{region 'Documentation'}
(*!
<summary>Checks results and isolated findings before allowing the script to advance.</summary>
*)
{endregion}
METHOD PROTECTED ProcessAssertions
VAR_INPUT
    Enable : BOOL; //! Phase permission supplied by the owning Test Case; FALSE does not authorize progression, while observation may continue.
END_VAR
VAR
    Evaluate : BOOL;
    FindingIndex : UINT;
    DetailsMatch : BOOL;
    FindingMatches : BOOL;
    ExpectedMessage : STRING(GVL_Constants.MessageLength);
END_VAR
FFirstCycleGate(Enable := Enable AND FGateObservationReady,
    State := State,
    IN := FGateMatches);
Evaluate := Enable AND FObservationReady;
FIsNaNResult(Enable := Evaluate,
    State := State,
    IN := FIsNaNSubject.Result = FExpectedIsNaN);
FIsFiniteResult(Enable := Evaluate,
    State := State,
    IN := FIsFiniteSubject.Result = FExpectedIsFinite);
FIsInfiniteResult(Enable := Evaluate,
    State := State,
    IN := FIsInfiniteSubject.Result = FExpectedIsInfinite);
DetailsMatch := TRUE;
FindingIndex := 1;
IF Evaluate THEN
    IF FFindingIsNaN <> E_Result.NotEvaluated THEN
        ExpectedMessage := CONCAT('Assertion failed: expected NaN. Actual = ',
            CreateAssertionTextValue_LReal(Value := FValue.Value));
        ExpectedMessage := CONCAT(ExpectedMessage, '.');
        FindingMatches := IsFindingValid(Index := FindingIndex,
            ExpectedName := FIsNaNSubject.Name,
            ExpectedResult := FFindingIsNaN,
            ExpectedMessage := ExpectedMessage);
        DetailsMatch := DetailsMatch AND FindingMatches;
        FindingIndex := FindingIndex + 1;
    END_IF;
    IF FFindingIsFinite <> E_Result.NotEvaluated THEN
        ExpectedMessage := CONCAT('Assertion failed: expected a finite value. Actual = ',
            CreateAssertionTextValue_LReal(Value := FValue.Value));
        ExpectedMessage := CONCAT(ExpectedMessage, '.');
        FindingMatches := IsFindingValid(Index := FindingIndex,
            ExpectedName := FIsFiniteSubject.Name,
            ExpectedResult := FFindingIsFinite,
            ExpectedMessage := ExpectedMessage);
        DetailsMatch := DetailsMatch AND FindingMatches;
        FindingIndex := FindingIndex + 1;
    END_IF;
    IF FFindingIsInfinite <> E_Result.NotEvaluated THEN
        ExpectedMessage := CONCAT('Assertion failed: expected positive or negative infinity. Actual = ',
            CreateAssertionTextValue_LReal(Value := FValue.Value));
        ExpectedMessage := CONCAT(ExpectedMessage, '.');
        FindingMatches := IsFindingValid(Index := FindingIndex,
            ExpectedName := FIsInfiniteSubject.Name,
            ExpectedResult := FFindingIsInfinite,
            ExpectedMessage := ExpectedMessage);
        DetailsMatch := DetailsMatch AND FindingMatches;
        FindingIndex := FindingIndex + 1;
    END_IF;
END_IF;
FCaptureIntegrity(Enable := Evaluate,
    State := State,
    IN := (FCaptureStatus.SequenceId = UINT_TO_UDINT(FindingIndex - 1))
        AND (FCaptureStatus.LostEventCount = 0)
        AND (FCaptureFifo.ElementCount = FindingIndex - 1));
FFindingDetails(Enable := Evaluate,
    State := State,
    IN := DetailsMatch);
IF Evaluate THEN
    FChecked := TRUE;
END_IF;
END_METHOD

{region 'Documentation'}
(*!
<summary>No Preparation phase is required.</summary>
*)
{endregion}
METHOD PROTECTED ProcessPreparations
VAR_INPUT
    // SA0033: Required hook; no Preparation phase.
    {attribute 'analysis' := '-33'}
    Enable : BOOL; //! Phase permission supplied by the owning Test Case; FALSE does not authorize progression, while observation may continue.
END_VAR
END_METHOD

{region 'Documentation'}
(*!
<summary>Restarts the row script and resets outer verdicts.</summary>
*)
{endregion}
METHOD PROTECTED ProcessReset
FFirstCycleGate.Reset();
FFirstCyclePending := FALSE;
FGateObservationReady := FALSE;
FGateMatches := FALSE;
FRow := RowQuietNaN;
FRowPrepared := FALSE;
FRepeatChecked := FALSE;
FChecked := FALSE;
FObservationReady := FALSE;
FIsNaNResult.Reset();
FIsFiniteResult.Reset();
FIsInfiniteResult.Reset();
FCaptureIntegrity.Reset();
FFindingDetails.Reset();
CompleteReset();
END_METHOD

{region 'Documentation'}
(*!
<summary>Prepares, checks and repeats each row over separate PLC cycles.</summary>
*)
{endregion}
METHOD PROTECTED ProcessTests
VAR_INPUT
    Enable : BOOL; //! Phase permission supplied by the owning Test Case; FALSE does not authorize progression, while observation may continue.
END_VAR
IF NOT Enable THEN
    RETURN;
END_IF;

FGateObservationReady := FALSE;
IF FChecked THEN
    FChecked := FALSE;
    FObservationReady := FALSE;
    IF FRepeatChecked THEN
        IF FRow = LastRow THEN
            CompleteTests();
            RETURN;
        END_IF;
        FRow := FRow + 1;
        FRowPrepared := FALSE;
        FRepeatChecked := FALSE;
    ELSE
        FRepeatChecked := TRUE;
    END_IF;
END_IF;

IF NOT FRowPrepared THEN
    SelectRow();
    FCapture.Reset();
    IF NOT FPreserveResults THEN
        ResetSubjects();
    END_IF;
    CallSubjects(Enable := FALSE);
    FRowPrepared := TRUE;
    FFirstCyclePending := TRUE;
ELSIF FFirstCyclePending THEN
    CallSubjects(Enable := FSubjectEnable);
    FFirstCyclePending := FALSE;
    FGateMatches := (FIsNaNSubject.Result = E_Result.NotEvaluated)
        AND (FIsFiniteSubject.Result = E_Result.NotEvaluated)
        AND (FIsInfiniteSubject.Result = E_Result.NotEvaluated)
        AND (FCaptureStatus.SequenceId = 0);
    FGateObservationReady := NOT FPreserveResults;
ELSE
    CallSubjects(Enable := FSubjectEnable);
    FObservationReady := TRUE;
END_IF;
END_METHOD

{region 'Documentation'}
(*!
<summary>Queues normal subject resets; CallSubjects consumes them.</summary>
*)
{endregion}
METHOD PRIVATE ResetSubjects
FIsNaNSubject.Reset();
FIsFiniteSubject.Reset();
FIsInfiniteSubject.Reset();
END_METHOD

{region 'Documentation'}
(*!
<summary>Supplies literal expectations; only named hold/escalation rows preserve subjects.</summary>
*)
{endregion}
METHOD PRIVATE SelectRow
FPreserveResults := FALSE;
FSubjectEnable := TRUE;

CASE FRow OF
    RowQuietNaN:
        FValue.Bits := QuietNaNBits;
        FExpectedIsNaN := E_Result.Passed;
        FFindingIsNaN := E_Result.NotEvaluated;
        FExpectedIsFinite := E_Result.Failed;
        FFindingIsFinite := E_Result.Failed;
        FExpectedIsInfinite := E_Result.Failed;
        FFindingIsInfinite := E_Result.Failed;
    RowSignalingNaN:
        FValue.Bits := SignalingNaNBits;
        FExpectedIsNaN := E_Result.Passed;
        FFindingIsNaN := E_Result.NotEvaluated;
        FExpectedIsFinite := E_Result.Failed;
        FFindingIsFinite := E_Result.Failed;
        FExpectedIsInfinite := E_Result.Failed;
        FFindingIsInfinite := E_Result.Failed;
    RowPositiveInfinity:
        FValue.Bits := PositiveInfinityBits;
        FExpectedIsNaN := E_Result.Failed;
        FFindingIsNaN := E_Result.Failed;
        FExpectedIsFinite := E_Result.Failed;
        FFindingIsFinite := E_Result.Failed;
        FExpectedIsInfinite := E_Result.Passed;
        FFindingIsInfinite := E_Result.NotEvaluated;
    RowNegativeInfinity:
        FValue.Bits := NegativeInfinityBits;
        FExpectedIsNaN := E_Result.Failed;
        FFindingIsNaN := E_Result.Failed;
        FExpectedIsFinite := E_Result.Failed;
        FFindingIsFinite := E_Result.Failed;
        FExpectedIsInfinite := E_Result.Passed;
        FFindingIsInfinite := E_Result.NotEvaluated;
    RowPositiveZero:
        FValue.Bits := PositiveZeroBits;
        FExpectedIsNaN := E_Result.Failed;
        FFindingIsNaN := E_Result.Failed;
        FExpectedIsFinite := E_Result.Passed;
        FFindingIsFinite := E_Result.NotEvaluated;
        FExpectedIsInfinite := E_Result.Failed;
        FFindingIsInfinite := E_Result.Failed;
    RowNegativeZero:
        FValue.Bits := NegativeZeroBits;
        FExpectedIsNaN := E_Result.Failed;
        FFindingIsNaN := E_Result.Failed;
        FExpectedIsFinite := E_Result.Passed;
        FFindingIsFinite := E_Result.NotEvaluated;
        FExpectedIsInfinite := E_Result.Failed;
        FFindingIsInfinite := E_Result.Failed;
    RowPositiveSubnormal:
        FValue.Bits := PositiveSubnormalBits;
        FExpectedIsNaN := E_Result.Failed;
        FFindingIsNaN := E_Result.Failed;
        FExpectedIsFinite := E_Result.Passed;
        FFindingIsFinite := E_Result.NotEvaluated;
        FExpectedIsInfinite := E_Result.Failed;
        FFindingIsInfinite := E_Result.Failed;
    RowNegativeSubnormal:
        FValue.Bits := NegativeSubnormalBits;
        FExpectedIsNaN := E_Result.Failed;
        FFindingIsNaN := E_Result.Failed;
        FExpectedIsFinite := E_Result.Passed;
        FFindingIsFinite := E_Result.NotEvaluated;
        FExpectedIsInfinite := E_Result.Failed;
        FFindingIsInfinite := E_Result.Failed;
    RowOrdinaryFinite:
        FValue.Bits := OrdinaryFiniteBits;
        FExpectedIsNaN := E_Result.Failed;
        FFindingIsNaN := E_Result.Failed;
        FExpectedIsFinite := E_Result.Passed;
        FFindingIsFinite := E_Result.NotEvaluated;
        FExpectedIsInfinite := E_Result.Failed;
        FFindingIsInfinite := E_Result.Failed;
    RowMaximumFinite:
        FValue.Bits := MaximumFiniteBits;
        FExpectedIsNaN := E_Result.Failed;
        FFindingIsNaN := E_Result.Failed;
        FExpectedIsFinite := E_Result.Passed;
        FFindingIsFinite := E_Result.NotEvaluated;
        FExpectedIsInfinite := E_Result.Failed;
        FFindingIsInfinite := E_Result.Failed;
    RowHoldResults:
        FValue.Bits := QuietNaNBits;
        FPreserveResults := TRUE;
        FExpectedIsNaN := E_Result.Failed;
        FFindingIsNaN := E_Result.NotEvaluated;
        FExpectedIsFinite := E_Result.Failed;
        FFindingIsFinite := E_Result.Failed;
        FExpectedIsInfinite := E_Result.Failed;
        FFindingIsInfinite := E_Result.NotEvaluated;
    RowDisabledHold:
        FValue.Bits := PositiveInfinityBits;
        FSubjectEnable := FALSE;
        FPreserveResults := TRUE;
        FExpectedIsNaN := E_Result.Failed;
        FFindingIsNaN := E_Result.NotEvaluated;
        FExpectedIsFinite := E_Result.Failed;
        FFindingIsFinite := E_Result.NotEvaluated;
        FExpectedIsInfinite := E_Result.Failed;
        FFindingIsInfinite := E_Result.NotEvaluated;
ELSE
    Error(Message := 'Unknown classification selftest row.');
END_CASE;
END_METHOD

END_FUNCTION_BLOCK

// ---- Framework/Assertions/POU/BasicTypes/LReal/AssertIsNaN_LReal.TcPOU
{region 'Documentation'}
(*!
<summary>Checks that IN is NaN.</summary>
<description>

NaN and either infinity are legitimate checked data, not configuration errors.
Classification mismatch reports Failed. Bit-based classification does not perform an ordered
floating-point comparison.

Numeric diagnostics use the formatter's default six significant digits; rounding affects
the message only, not the comparison.

</description>
*)
{endregion}
FUNCTION_BLOCK AssertIsNaN_LReal EXTENDS AssertionBase
VAR_INPUT
    IN : LREAL; //! Value to classify; NaN and both infinities are valid inputs.
END_VAR

SUPER^();

{region 'Documentation'}
(*!
<summary>Classifies the bit representation without floating-point arithmetic.</summary>
*)
{endregion}
METHOD PROTECTED Assert
VAR
    Representation : AssertionLRealRepresentation;
    Message : STRING(GVL_Constants.MessageLength);
END_VAR
VAR CONSTANT
    ExponentMask : LWORD := LWORD#16#7FF0000000000000;
    FractionMask : LWORD := LWORD#16#000FFFFFFFFFFFFF;
END_VAR
IF NOT EvaluationActive THEN
    RETURN;
END_IF;

IF Result = E_Result.Error THEN
    RETURN;
END_IF;

IF Result = E_Result.Failed THEN
    RETURN;
END_IF;

Representation.Value := IN;
IF ((Representation.Bits AND ExponentMask) <> ExponentMask)
    OR ((Representation.Bits AND FractionMask) = 0) THEN
    Message := CONCAT('Assertion failed: expected NaN. Actual = ',
        CreateAssertionTextValue_LReal(Value := IN));
    Message := CONCAT(Message, '.');
    Fail(Message := Message);
    RETURN;
END_IF;

Pass();
END_METHOD

END_FUNCTION_BLOCK

// ---- Framework/Assertions/POU/BasicTypes/LReal/AssertIsFinite_LReal.TcPOU
{region 'Documentation'}
(*!
<summary>Checks that IN is a finite value.</summary>
<description>

NaN and either infinity are legitimate checked data, not configuration errors.
Classification mismatch reports Failed. Bit-based classification does not perform an ordered
floating-point comparison.

Numeric diagnostics use the formatter's default six significant digits; rounding affects
the message only, not the comparison.

</description>
*)
{endregion}
FUNCTION_BLOCK AssertIsFinite_LReal EXTENDS AssertionBase
VAR_INPUT
    IN : LREAL; //! Value to classify; NaN and both infinities are valid inputs.
END_VAR

SUPER^();

{region 'Documentation'}
(*!
<summary>Classifies the bit representation without floating-point arithmetic.</summary>
*)
{endregion}
METHOD PROTECTED Assert
VAR
    Representation : AssertionLRealRepresentation;
    Message : STRING(GVL_Constants.MessageLength);
END_VAR
VAR CONSTANT
    ExponentMask : LWORD := LWORD#16#7FF0000000000000;
END_VAR
IF NOT EvaluationActive THEN
    RETURN;
END_IF;

IF Result = E_Result.Error THEN
    RETURN;
END_IF;

IF Result = E_Result.Failed THEN
    RETURN;
END_IF;

Representation.Value := IN;
IF (Representation.Bits AND ExponentMask) = ExponentMask THEN
    Message := CONCAT('Assertion failed: expected a finite value. Actual = ',
        CreateAssertionTextValue_LReal(Value := IN));
    Message := CONCAT(Message, '.');
    Fail(Message := Message);
    RETURN;
END_IF;

Pass();
END_METHOD

END_FUNCTION_BLOCK

// ---- Framework/Assertions/POU/BasicTypes/LReal/AssertIsInfinite_LReal.TcPOU
{region 'Documentation'}
(*!
<summary>Checks that IN is positive or negative infinity.</summary>
<description>

NaN and either infinity are legitimate checked data, not configuration errors.
Classification mismatch reports Failed. Bit-based classification does not perform an ordered
floating-point comparison.

Numeric diagnostics use the formatter's default six significant digits; rounding affects
the message only, not the comparison.

</description>
*)
{endregion}
FUNCTION_BLOCK AssertIsInfinite_LReal EXTENDS AssertionBase
VAR_INPUT
    IN : LREAL; //! Value to classify; NaN and both infinities are valid inputs.
END_VAR

SUPER^();

{region 'Documentation'}
(*!
<summary>Classifies the bit representation without floating-point arithmetic.</summary>
*)
{endregion}
METHOD PROTECTED Assert
VAR
    Representation : AssertionLRealRepresentation;
    Message : STRING(GVL_Constants.MessageLength);
END_VAR
VAR CONSTANT
    ExponentMask : LWORD := LWORD#16#7FF0000000000000;
    FractionMask : LWORD := LWORD#16#000FFFFFFFFFFFFF;
END_VAR
IF NOT EvaluationActive THEN
    RETURN;
END_IF;

IF Result = E_Result.Error THEN
    RETURN;
END_IF;

IF Result = E_Result.Failed THEN
    RETURN;
END_IF;

Representation.Value := IN;
IF ((Representation.Bits AND ExponentMask) <> ExponentMask)
    OR ((Representation.Bits AND FractionMask) <> 0) THEN
    Message := CONCAT('Assertion failed: expected positive or negative infinity. Actual = ',
        CreateAssertionTextValue_LReal(Value := IN));
    Message := CONCAT(Message, '.');
    Fail(Message := Message);
    RETURN;
END_IF;

Pass();
END_METHOD

END_FUNCTION_BLOCK

// ---- SelfTests/TestCases/TestSuite_AssertionFloatingPoint/Test_AssertionArrayClassification_LReal.TcPOU
{region 'Documentation'}
(*!
<summary>Checks LREAL array classification with literal expected results and isolated findings.</summary>
<description>
Each named row selects checked data and independent expected outcomes.
SelectRow does not derive expectations from the production classification algorithm.
A disabled preparation call consumes subject reset requests before evaluation.
The first enabled call is checked, then repeated on the next cycle to verify no duplicate finding.
Only outer Assertions contribute to the Test Case; deliberate subject failures stay in the local capture.
Named preservation rows check Failed-to-Error escalation and held Error; other rows reset subjects.
Special values are supplied by integer bit patterns, never exceptional floating-point arithmetic.
</description>
*)
{endregion}
FUNCTION_BLOCK Test_AssertionArrayClassification_LReal EXTENDS TestCaseBase
VAR
    FAllElementsFiniteSubject : AssertArrayAllElementsFinite_LReal;
    FAllElementsFiniteResult : AssertTrue;
    FExpectedAllElementsFinite : E_Result;
    FFindingAllElementsFinite : E_Result;
    FContainsNonFiniteSubject : AssertArrayContainsNonFinite_LReal;
    FContainsNonFiniteResult : AssertTrue;
    FExpectedContainsNonFinite : E_Result;
    FFindingContainsNonFinite : E_Result;
    FContainsNaNSubject : AssertArrayContainsNaN_LReal;
    FContainsNaNResult : AssertTrue;
    FExpectedContainsNaN : E_Result;
    FFindingContainsNaN : E_Result;
    FHasNoNaNSubject : AssertArrayHasNoNaN_LReal;
    FHasNoNaNResult : AssertTrue;
    FExpectedHasNoNaN : E_Result;
    FFindingHasNoNaN : E_Result;
    FContainsInfinitySubject : AssertArrayContainsInfinity_LReal;
    FContainsInfinityResult : AssertTrue;
    FExpectedContainsInfinity : E_Result;
    FFindingContainsInfinity : E_Result;
    FHasNoInfinitySubject : AssertArrayHasNoInfinity_LReal;
    FHasNoInfinityResult : AssertTrue;
    FExpectedHasNoInfinity : E_Result;
    FFindingHasNoInfinity : E_Result;
    FCaptureIntegrity : AssertTrue;
    FFindingDetails : AssertTrue;
    FCapture : EventBuffer;
    FEvents : ARRAY[1..CaptureLength] OF ST_Event;
    FCaptureFifo : ST_FifoStatus;
    FCaptureStatus : ST_EventBufferStatus;
    FValues : ARRAY[-2..2] OF LREAL;
    FStartIndex : DINT;
    FLength : USINT;
    FExpectedIndex : DINT;
    FExpectedInfinityIndex : DINT;
    FQuietNaN : FloatingPointBits_LReal;
    FSignalingNaN : FloatingPointBits_LReal;
    FPositiveInfinity : FloatingPointBits_LReal;
    FNegativeInfinity : FloatingPointBits_LReal;
    FPositiveZero : FloatingPointBits_LReal;
    FNegativeZero : FloatingPointBits_LReal;
    FPositiveSubnormal : FloatingPointBits_LReal;
    FNegativeSubnormal : FloatingPointBits_LReal;
    FOrdinaryFinite : FloatingPointBits_LReal;
    FMaximumFinite : FloatingPointBits_LReal;
    FRow : UINT;
    FRowPrepared : BOOL;
    FRepeatChecked : BOOL;
    FChecked : BOOL;
    FObservationReady : BOOL;
    FPreserveResults : BOOL;
    FSubjectEnable : BOOL;
    FSetupValid : BOOL;
END_VAR
VAR CONSTANT
    CaptureLength : UINT := 16;
    QuietNaNBits : LWORD := LWORD#16#7FF8000000000000;
    SignalingNaNBits : LWORD := LWORD#16#7FF0000000000001;
    PositiveInfinityBits : LWORD := LWORD#16#7FF0000000000000;
    NegativeInfinityBits : LWORD := LWORD#16#FFF0000000000000;
    PositiveZeroBits : LWORD := LWORD#16#0000000000000000;
    NegativeZeroBits : LWORD := LWORD#16#8000000000000000;
    PositiveSubnormalBits : LWORD := LWORD#16#0000000000000001;
    NegativeSubnormalBits : LWORD := LWORD#16#8000000000000001;
    OrdinaryFiniteBits : LWORD := LWORD#16#3FF0000000000000;
    MaximumFiniteBits : LWORD := LWORD#16#7FEFFFFFFFFFFFFF;
    RowFiniteValues : UINT := 1;
    RowNaNFirst : UINT := 2;
    RowSignalingNaNMiddle : UINT := 3;
    RowNaNLast : UINT := 4;
    RowInfinityFirst : UINT := 5;
    RowInfinityMiddle : UINT := 6;
    RowInfinityLast : UINT := 7;
    RowMixedSpecials : UINT := 8;
    RowOutsideSelection : UINT := 9;
    RowSingleLastElement : UINT := 10;
    RowInvalidAfterFailed : UINT := 11;
    RowErrorRemainsHeld : UINT := 12;
    RowStartBelowBounds : UINT := 13;
    RowStartAboveBounds : UINT := 14;
    RowEndAboveBounds : UINT := 15;
    RowLargeStart : UINT := 16;
    RowZeroLength : UINT := 17;
    RowResetRecovers : UINT := 18;
    LastRow : UINT := RowResetRecovers;
END_VAR

SUPER^();

{region 'Documentation'}
(*!
<summary>Collects verdicts, excluding deliberate subject findings.</summary>
*)
{endregion}
METHOD PROTECTED AggregateResults
VAR_INPUT
    Aggregator : I_ResultAggregator; //! Borrowed result sink owned by the outer Test Case; add this test's checking Assertions without resetting or retaining the sink.
END_VAR
Aggregator.AddProvider(Provider := FAllElementsFiniteResult);
Aggregator.AddProvider(Provider := FContainsNonFiniteResult);
Aggregator.AddProvider(Provider := FContainsNaNResult);
Aggregator.AddProvider(Provider := FHasNoNaNResult);
Aggregator.AddProvider(Provider := FContainsInfinityResult);
Aggregator.AddProvider(Provider := FHasNoInfinityResult);
Aggregator.AddProvider(Provider := FCaptureIntegrity);
Aggregator.AddProvider(Provider := FFindingDetails);
END_METHOD

{region 'Documentation'}
(*!
<summary>Calls each concrete production subject with the selected data.</summary>
*)
{endregion}
METHOD PRIVATE CallSubjects
VAR_INPUT
    Enable : BOOL; //! Observation-enable input forwarded to the controlled Assertion subjects for this call.
END_VAR
FAllElementsFiniteSubject(Enable := Enable,
    State := E_State.Running,
    StartIndex := FStartIndex,
    Length := FLength,
    IN := FValues);
FContainsNonFiniteSubject(Enable := Enable,
    State := E_State.Running,
    StartIndex := FStartIndex,
    Length := FLength,
    IN := FValues);
FContainsNaNSubject(Enable := Enable,
    State := E_State.Running,
    StartIndex := FStartIndex,
    Length := FLength,
    IN := FValues);
FHasNoNaNSubject(Enable := Enable,
    State := E_State.Running,
    StartIndex := FStartIndex,
    Length := FLength,
    IN := FValues);
FContainsInfinitySubject(Enable := Enable,
    State := E_State.Running,
    StartIndex := FStartIndex,
    Length := FLength,
    IN := FValues);
FHasNoInfinitySubject(Enable := Enable,
    State := E_State.Running,
    StartIndex := FStartIndex,
    Length := FLength,
    IN := FValues);
END_METHOD

{region 'Documentation'}
(*!
<summary>Rejects incomplete subject or verdict setup.</summary>
*)
{endregion}
METHOD PROTECTED CheckInitialization : BOOL //! TRUE when the inherited initialization check and this concrete fixture check both accept the setup.
CheckInitialization := SUPER^.CheckInitialization();
IF NOT CheckInitialization THEN
    RETURN;
END_IF;
CheckInitialization := FSetupValid
    AND FAllElementsFiniteResult.IsInitialized
    AND FContainsNonFiniteResult.IsInitialized
    AND FContainsNaNResult.IsInitialized
    AND FHasNoNaNResult.IsInitialized
    AND FContainsInfinityResult.IsInitialized
    AND FHasNoInfinityResult.IsInitialized
    AND FCaptureIntegrity.IsInitialized
    AND FFindingDetails.IsInitialized;
END_METHOD

{region 'Documentation'}
(*!
<summary>Initializes isolated subjects and the outer verdict Assertions.</summary>
*)
{endregion}
METHOD PROTECTED Configure
VAR
    Initialized : BOOL;
END_VAR
FPreparationStateCount := 0;
FTestStateCount := 1;
FQuietNaN.Bits := QuietNaNBits;
FSignalingNaN.Bits := SignalingNaNBits;
FPositiveInfinity.Bits := PositiveInfinityBits;
FNegativeInfinity.Bits := NegativeInfinityBits;
FPositiveZero.Bits := PositiveZeroBits;
FNegativeZero.Bits := NegativeZeroBits;
FPositiveSubnormal.Bits := PositiveSubnormalBits;
FNegativeSubnormal.Bits := NegativeSubnormalBits;
FOrdinaryFinite.Bits := OrdinaryFiniteBits;
FMaximumFinite.Bits := MaximumFiniteBits;
FSetupValid := FCapture.Initialize(Buffer := FEvents,
    FifoControl := FCaptureFifo,
    Status := FCaptureStatus);
FAllElementsFiniteResult.Initialize(Parent := THIS^,
    AssertionName := 'AllElementsFiniteResult');
FContainsNonFiniteResult.Initialize(Parent := THIS^,
    AssertionName := 'ContainsNonFiniteResult');
FContainsNaNResult.Initialize(Parent := THIS^,
    AssertionName := 'ContainsNaNResult');
FHasNoNaNResult.Initialize(Parent := THIS^,
    AssertionName := 'HasNoNaNResult');
FContainsInfinityResult.Initialize(Parent := THIS^,
    AssertionName := 'ContainsInfinityResult');
FHasNoInfinityResult.Initialize(Parent := THIS^,
    AssertionName := 'HasNoInfinityResult');
FCaptureIntegrity.Initialize(Parent := THIS^,
    AssertionName := 'CaptureIntegrity');
FFindingDetails.Initialize(Parent := THIS^,
    AssertionName := 'FindingDetails');
FAllElementsFiniteSubject.BindPublisher(Publisher := FCapture);
Initialized := FAllElementsFiniteSubject.Initialize(Parent := THIS^,
    AssertionName := 'AllElementsFiniteSubject');
FSetupValid := FSetupValid AND Initialized;
FContainsNonFiniteSubject.BindPublisher(Publisher := FCapture);
Initialized := FContainsNonFiniteSubject.Initialize(Parent := THIS^,
    AssertionName := 'ContainsNonFiniteSubject');
FSetupValid := FSetupValid AND Initialized;
FContainsNaNSubject.BindPublisher(Publisher := FCapture);
Initialized := FContainsNaNSubject.Initialize(Parent := THIS^,
    AssertionName := 'ContainsNaNSubject');
FSetupValid := FSetupValid AND Initialized;
FHasNoNaNSubject.BindPublisher(Publisher := FCapture);
Initialized := FHasNoNaNSubject.Initialize(Parent := THIS^,
    AssertionName := 'HasNoNaNSubject');
FSetupValid := FSetupValid AND Initialized;
FContainsInfinitySubject.BindPublisher(Publisher := FCapture);
Initialized := FContainsInfinitySubject.Initialize(Parent := THIS^,
    AssertionName := 'ContainsInfinitySubject');
FSetupValid := FSetupValid AND Initialized;
FHasNoInfinitySubject.BindPublisher(Publisher := FCapture);
Initialized := FHasNoInfinitySubject.Initialize(Parent := THIS^,
    AssertionName := 'HasNoInfinitySubject');
FSetupValid := FSetupValid AND Initialized;
END_METHOD

{region 'Documentation'}
(*!
<summary>Checks ordered capture metadata and meaningful diagnostic text.</summary>
*)
{endregion}
METHOD PRIVATE IsFindingValid : BOOL //! TRUE when the selected captured finding satisfies the scenario metadata and diagnostic checks.
VAR_INPUT
    Index : UINT; //! One-based index in the retained isolated event capture.
    ExpectedName : STRING(GVL_Constants.NameLength); //! Independently authored Assertion name expected in the selected finding.
    ExpectedResult : E_Result; //! Independently authored finding result.
    ExpectedMessage : STRING(GVL_Constants.MessageLength); //! Exact diagnostic text expected in the selected finding.
END_VAR
IsFindingValid := (FEvents[Index].SequenceId = UINT_TO_UDINT(Index))
    AND (FEvents[Index].Name = ExpectedName)
    AND (FEvents[Index].OwnerScope = E_OwnerScope.Assertion)
    AND (FEvents[Index].EventType = E_EventType.Result)
    AND (FEvents[Index].State = E_State.Running)
    AND (FEvents[Index].Result = ExpectedResult)
    AND (FEvents[Index].Message <> '')
    AND (FEvents[Index].Message = ExpectedMessage);
END_METHOD

{region 'Documentation'}
(*!
<summary>No asynchronous cleanup is needed.</summary>
*)
{endregion}
METHOD PROTECTED ProcessAbort
VAR_INPUT
    Enable : BOOL; //! Phase permission supplied by the owning Test Case; FALSE does not authorize progression, while observation may continue.
END_VAR
IF Enable THEN
    CompleteAbort();
END_IF;
END_METHOD

{region 'Documentation'}
(*!
<summary>Checks results and isolated findings before allowing the script to advance.</summary>
*)
{endregion}
METHOD PROTECTED ProcessAssertions
VAR_INPUT
    Enable : BOOL; //! Phase permission supplied by the owning Test Case; FALSE does not authorize progression, while observation may continue.
END_VAR
VAR
    Evaluate : BOOL;
    FindingIndex : UINT;
    DetailsMatch : BOOL;
    FindingMatches : BOOL;
    ExpectedMessage : STRING(GVL_Constants.MessageLength);
END_VAR
Evaluate := Enable AND FObservationReady;
FAllElementsFiniteResult(Enable := Evaluate,
    State := State,
    IN := FAllElementsFiniteSubject.Result = FExpectedAllElementsFinite);
FContainsNonFiniteResult(Enable := Evaluate,
    State := State,
    IN := FContainsNonFiniteSubject.Result = FExpectedContainsNonFinite);
FContainsNaNResult(Enable := Evaluate,
    State := State,
    IN := FContainsNaNSubject.Result = FExpectedContainsNaN);
FHasNoNaNResult(Enable := Evaluate,
    State := State,
    IN := FHasNoNaNSubject.Result = FExpectedHasNoNaN);
FContainsInfinityResult(Enable := Evaluate,
    State := State,
    IN := FContainsInfinitySubject.Result = FExpectedContainsInfinity);
FHasNoInfinityResult(Enable := Evaluate,
    State := State,
    IN := FHasNoInfinitySubject.Result = FExpectedHasNoInfinity);
DetailsMatch := TRUE;
FindingIndex := 1;
IF Evaluate THEN
    IF FFindingAllElementsFinite <> E_Result.NotEvaluated THEN
        IF FFindingAllElementsFinite = E_Result.Error THEN
            ExpectedMessage := CONCAT('Assertion error: array range is invalid. StartIndex = ',
                DINT_TO_STRING(FStartIndex));
            ExpectedMessage := CONCAT(ExpectedMessage, ', Length = ');
            ExpectedMessage := CONCAT(ExpectedMessage, USINT_TO_STRING(FLength));
            ExpectedMessage := CONCAT(ExpectedMessage, '.');
        ELSE
            ExpectedMessage := 'Assertion failed: array range contains a non-finite value.';
            ExpectedMessage := CONCAT(ExpectedMessage, ' Actual[');
            ExpectedMessage := CONCAT(ExpectedMessage, DINT_TO_STRING(FExpectedIndex));
            ExpectedMessage := CONCAT(ExpectedMessage, '] = ');
            ExpectedMessage := CONCAT(ExpectedMessage, CreateAssertionTextValue_LReal(Value := FValues[FExpectedIndex]));
            ExpectedMessage := CONCAT(ExpectedMessage, ', Range = [');
            ExpectedMessage := CONCAT(ExpectedMessage, DINT_TO_STRING(FStartIndex));
            ExpectedMessage := CONCAT(ExpectedMessage, '..');
            ExpectedMessage := CONCAT(ExpectedMessage, LINT_TO_STRING(DINT_TO_LINT(FStartIndex) + USINT_TO_LINT(FLength) - 1));
            ExpectedMessage := CONCAT(ExpectedMessage, '].');
        END_IF;
        FindingMatches := IsFindingValid(Index := FindingIndex,
            ExpectedName := FAllElementsFiniteSubject.Name,
            ExpectedResult := FFindingAllElementsFinite,
            ExpectedMessage := ExpectedMessage);
        DetailsMatch := DetailsMatch AND FindingMatches;
        FindingIndex := FindingIndex + 1;
    END_IF;
    IF FFindingContainsNonFinite <> E_Result.NotEvaluated THEN
        IF FFindingContainsNonFinite = E_Result.Error THEN
            ExpectedMessage := CONCAT('Assertion error: array range is invalid. StartIndex = ',
                DINT_TO_STRING(FStartIndex));
            ExpectedMessage := CONCAT(ExpectedMessage, ', Length = ');
            ExpectedMessage := CONCAT(ExpectedMessage, USINT_TO_STRING(FLength));
            ExpectedMessage := CONCAT(ExpectedMessage, '.');
        ELSE
            ExpectedMessage := 'Assertion failed: array range contains no non-finite value.';
            ExpectedMessage := CONCAT(ExpectedMessage, ', Range = [');
            ExpectedMessage := CONCAT(ExpectedMessage, DINT_TO_STRING(FStartIndex));
            ExpectedMessage := CONCAT(ExpectedMessage, '..');
            ExpectedMessage := CONCAT(ExpectedMessage, LINT_TO_STRING(DINT_TO_LINT(FStartIndex) + USINT_TO_LINT(FLength) - 1));
            ExpectedMessage := CONCAT(ExpectedMessage, '].');
        END_IF;
        FindingMatches := IsFindingValid(Index := FindingIndex,
            ExpectedName := FContainsNonFiniteSubject.Name,
            ExpectedResult := FFindingContainsNonFinite,
            ExpectedMessage := ExpectedMessage);
        DetailsMatch := DetailsMatch AND FindingMatches;
        FindingIndex := FindingIndex + 1;
    END_IF;
    IF FFindingContainsNaN <> E_Result.NotEvaluated THEN
        IF FFindingContainsNaN = E_Result.Error THEN
            ExpectedMessage := CONCAT('Assertion error: array range is invalid. StartIndex = ',
                DINT_TO_STRING(FStartIndex));
            ExpectedMessage := CONCAT(ExpectedMessage, ', Length = ');
            ExpectedMessage := CONCAT(ExpectedMessage, USINT_TO_STRING(FLength));
            ExpectedMessage := CONCAT(ExpectedMessage, '.');
        ELSE
            ExpectedMessage := 'Assertion failed: array range contains no NaN.';
            ExpectedMessage := CONCAT(ExpectedMessage, ', Range = [');
            ExpectedMessage := CONCAT(ExpectedMessage, DINT_TO_STRING(FStartIndex));
            ExpectedMessage := CONCAT(ExpectedMessage, '..');
            ExpectedMessage := CONCAT(ExpectedMessage, LINT_TO_STRING(DINT_TO_LINT(FStartIndex) + USINT_TO_LINT(FLength) - 1));
            ExpectedMessage := CONCAT(ExpectedMessage, '].');
        END_IF;
        FindingMatches := IsFindingValid(Index := FindingIndex,
            ExpectedName := FContainsNaNSubject.Name,
            ExpectedResult := FFindingContainsNaN,
            ExpectedMessage := ExpectedMessage);
        DetailsMatch := DetailsMatch AND FindingMatches;
        FindingIndex := FindingIndex + 1;
    END_IF;
    IF FFindingHasNoNaN <> E_Result.NotEvaluated THEN
        IF FFindingHasNoNaN = E_Result.Error THEN
            ExpectedMessage := CONCAT('Assertion error: array range is invalid. StartIndex = ',
                DINT_TO_STRING(FStartIndex));
            ExpectedMessage := CONCAT(ExpectedMessage, ', Length = ');
            ExpectedMessage := CONCAT(ExpectedMessage, USINT_TO_STRING(FLength));
            ExpectedMessage := CONCAT(ExpectedMessage, '.');
        ELSE
            ExpectedMessage := 'Assertion failed: array range contains NaN.';
            ExpectedMessage := CONCAT(ExpectedMessage, ' Actual[');
            ExpectedMessage := CONCAT(ExpectedMessage, DINT_TO_STRING(FExpectedIndex));
            ExpectedMessage := CONCAT(ExpectedMessage, '] = ');
            ExpectedMessage := CONCAT(ExpectedMessage, CreateAssertionTextValue_LReal(Value := FValues[FExpectedIndex]));
            ExpectedMessage := CONCAT(ExpectedMessage, ', Range = [');
            ExpectedMessage := CONCAT(ExpectedMessage, DINT_TO_STRING(FStartIndex));
            ExpectedMessage := CONCAT(ExpectedMessage, '..');
            ExpectedMessage := CONCAT(ExpectedMessage, LINT_TO_STRING(DINT_TO_LINT(FStartIndex) + USINT_TO_LINT(FLength) - 1));
            ExpectedMessage := CONCAT(ExpectedMessage, '].');
        END_IF;
        FindingMatches := IsFindingValid(Index := FindingIndex,
            ExpectedName := FHasNoNaNSubject.Name,
            ExpectedResult := FFindingHasNoNaN,
            ExpectedMessage := ExpectedMessage);
        DetailsMatch := DetailsMatch AND FindingMatches;
        FindingIndex := FindingIndex + 1;
    END_IF;
    IF FFindingContainsInfinity <> E_Result.NotEvaluated THEN
        IF FFindingContainsInfinity = E_Result.Error THEN
            ExpectedMessage := CONCAT('Assertion error: array range is invalid. StartIndex = ',
                DINT_TO_STRING(FStartIndex));
            ExpectedMessage := CONCAT(ExpectedMessage, ', Length = ');
            ExpectedMessage := CONCAT(ExpectedMessage, USINT_TO_STRING(FLength));
            ExpectedMessage := CONCAT(ExpectedMessage, '.');
        ELSE
            ExpectedMessage := 'Assertion failed: array range contains no infinity.';
            ExpectedMessage := CONCAT(ExpectedMessage, ', Range = [');
            ExpectedMessage := CONCAT(ExpectedMessage, DINT_TO_STRING(FStartIndex));
            ExpectedMessage := CONCAT(ExpectedMessage, '..');
            ExpectedMessage := CONCAT(ExpectedMessage, LINT_TO_STRING(DINT_TO_LINT(FStartIndex) + USINT_TO_LINT(FLength) - 1));
            ExpectedMessage := CONCAT(ExpectedMessage, '].');
        END_IF;
        FindingMatches := IsFindingValid(Index := FindingIndex,
            ExpectedName := FContainsInfinitySubject.Name,
            ExpectedResult := FFindingContainsInfinity,
            ExpectedMessage := ExpectedMessage);
        DetailsMatch := DetailsMatch AND FindingMatches;
        FindingIndex := FindingIndex + 1;
    END_IF;
    IF FFindingHasNoInfinity <> E_Result.NotEvaluated THEN
        IF FFindingHasNoInfinity = E_Result.Error THEN
            ExpectedMessage := CONCAT('Assertion error: array range is invalid. StartIndex = ',
                DINT_TO_STRING(FStartIndex));
            ExpectedMessage := CONCAT(ExpectedMessage, ', Length = ');
            ExpectedMessage := CONCAT(ExpectedMessage, USINT_TO_STRING(FLength));
            ExpectedMessage := CONCAT(ExpectedMessage, '.');
        ELSE
            ExpectedMessage := 'Assertion failed: array range contains infinity.';
            ExpectedMessage := CONCAT(ExpectedMessage, ' Actual[');
            ExpectedMessage := CONCAT(ExpectedMessage, DINT_TO_STRING(SEL(FRow = RowMixedSpecials, FExpectedIndex, FExpectedInfinityIndex)));
            ExpectedMessage := CONCAT(ExpectedMessage, '] = ');
            ExpectedMessage := CONCAT(ExpectedMessage, CreateAssertionTextValue_LReal(Value := FValues[SEL(FRow = RowMixedSpecials, FExpectedIndex, FExpectedInfinityIndex)]));
            ExpectedMessage := CONCAT(ExpectedMessage, ', Range = [');
            ExpectedMessage := CONCAT(ExpectedMessage, DINT_TO_STRING(FStartIndex));
            ExpectedMessage := CONCAT(ExpectedMessage, '..');
            ExpectedMessage := CONCAT(ExpectedMessage, LINT_TO_STRING(DINT_TO_LINT(FStartIndex) + USINT_TO_LINT(FLength) - 1));
            ExpectedMessage := CONCAT(ExpectedMessage, '].');
        END_IF;
        FindingMatches := IsFindingValid(Index := FindingIndex,
            ExpectedName := FHasNoInfinitySubject.Name,
            ExpectedResult := FFindingHasNoInfinity,
            ExpectedMessage := ExpectedMessage);
        DetailsMatch := DetailsMatch AND FindingMatches;
        FindingIndex := FindingIndex + 1;
    END_IF;
END_IF;
FCaptureIntegrity(Enable := Evaluate,
    State := State,
    IN := (FCaptureStatus.SequenceId = UINT_TO_UDINT(FindingIndex - 1))
        AND (FCaptureStatus.LostEventCount = 0)
        AND (FCaptureFifo.ElementCount = FindingIndex - 1));
FFindingDetails(Enable := Evaluate,
    State := State,
    IN := DetailsMatch);
IF Evaluate THEN
    FChecked := TRUE;
END_IF;
END_METHOD

{region 'Documentation'}
(*!
<summary>No Preparation phase is required.</summary>
*)
{endregion}
METHOD PROTECTED ProcessPreparations
VAR_INPUT
    // SA0033: Required hook; no Preparation phase.
    {attribute 'analysis' := '-33'}
    Enable : BOOL; //! Phase permission supplied by the owning Test Case; FALSE does not authorize progression, while observation may continue.
END_VAR
END_METHOD

{region 'Documentation'}
(*!
<summary>Restarts the row script and resets outer verdicts.</summary>
*)
{endregion}
METHOD PROTECTED ProcessReset
FRow := RowFiniteValues;
FRowPrepared := FALSE;
FRepeatChecked := FALSE;
FChecked := FALSE;
FObservationReady := FALSE;
FAllElementsFiniteResult.Reset();
FContainsNonFiniteResult.Reset();
FContainsNaNResult.Reset();
FHasNoNaNResult.Reset();
FContainsInfinityResult.Reset();
FHasNoInfinityResult.Reset();
FCaptureIntegrity.Reset();
FFindingDetails.Reset();
CompleteReset();
END_METHOD

{region 'Documentation'}
(*!
<summary>Prepares, checks and repeats each row over separate PLC cycles.</summary>
*)
{endregion}
METHOD PROTECTED ProcessTests
VAR_INPUT
    Enable : BOOL; //! Phase permission supplied by the owning Test Case; FALSE does not authorize progression, while observation may continue.
END_VAR
IF NOT Enable THEN
    RETURN;
END_IF;

IF FChecked THEN
    FChecked := FALSE;
    FObservationReady := FALSE;
    IF FRepeatChecked THEN
        IF FRow = LastRow THEN
            CompleteTests();
            RETURN;
        END_IF;
        FRow := FRow + 1;
        FRowPrepared := FALSE;
        FRepeatChecked := FALSE;
    ELSE
        FRepeatChecked := TRUE;
    END_IF;
END_IF;

IF NOT FRowPrepared THEN
    SelectRow();
    FCapture.Reset();
    IF NOT FPreserveResults THEN
        ResetSubjects();
    END_IF;
    CallSubjects(Enable := FALSE);
    FRowPrepared := TRUE;
ELSE
    CallSubjects(Enable := FSubjectEnable);
    FObservationReady := TRUE;
END_IF;
END_METHOD

{region 'Documentation'}
(*!
<summary>Queues normal subject resets; CallSubjects consumes them.</summary>
*)
{endregion}
METHOD PRIVATE ResetSubjects
FAllElementsFiniteSubject.Reset();
FContainsNonFiniteSubject.Reset();
FContainsNaNSubject.Reset();
FHasNoNaNSubject.Reset();
FContainsInfinitySubject.Reset();
FHasNoInfinitySubject.Reset();
END_METHOD

{region 'Documentation'}
(*!
<summary>Supplies literal expectations; only named hold/escalation rows preserve subjects.</summary>
*)
{endregion}
METHOD PRIVATE SelectRow
VAR
    Index : DINT;
END_VAR
FPreserveResults := FALSE;
FSubjectEnable := TRUE;
FStartIndex := -2;
FLength := 5;
FExpectedIndex := -2;
FExpectedInfinityIndex := -2;
FOR Index := -2 TO 2 DO
    FValues[Index] := FOrdinaryFinite.Value;
END_FOR;

CASE FRow OF
    RowFiniteValues:
        FValues[-2] := FPositiveZero.Value;
        FValues[-1] := FNegativeZero.Value;
        FValues[0] := FPositiveSubnormal.Value;
        FValues[1] := FNegativeSubnormal.Value;
        FValues[2] := FMaximumFinite.Value;
        FExpectedAllElementsFinite := E_Result.Passed;
        FFindingAllElementsFinite := E_Result.NotEvaluated;
        FExpectedContainsNonFinite := E_Result.Failed;
        FFindingContainsNonFinite := E_Result.Failed;
        FExpectedContainsNaN := E_Result.Failed;
        FFindingContainsNaN := E_Result.Failed;
        FExpectedHasNoNaN := E_Result.Passed;
        FFindingHasNoNaN := E_Result.NotEvaluated;
        FExpectedContainsInfinity := E_Result.Failed;
        FFindingContainsInfinity := E_Result.Failed;
        FExpectedHasNoInfinity := E_Result.Passed;
        FFindingHasNoInfinity := E_Result.NotEvaluated;
    RowNaNFirst:
        FValues[-2] := FQuietNaN.Value;
        FExpectedIndex := -2;
        FExpectedAllElementsFinite := E_Result.Failed;
        FFindingAllElementsFinite := E_Result.Failed;
        FExpectedContainsNonFinite := E_Result.Passed;
        FFindingContainsNonFinite := E_Result.NotEvaluated;
        FExpectedContainsNaN := E_Result.Passed;
        FFindingContainsNaN := E_Result.NotEvaluated;
        FExpectedHasNoNaN := E_Result.Failed;
        FFindingHasNoNaN := E_Result.Failed;
        FExpectedContainsInfinity := E_Result.Failed;
        FFindingContainsInfinity := E_Result.Failed;
        FExpectedHasNoInfinity := E_Result.Passed;
        FFindingHasNoInfinity := E_Result.NotEvaluated;
    RowSignalingNaNMiddle:
        FValues[0] := FSignalingNaN.Value;
        FExpectedIndex := 0;
        FExpectedAllElementsFinite := E_Result.Failed;
        FFindingAllElementsFinite := E_Result.Failed;
        FExpectedContainsNonFinite := E_Result.Passed;
        FFindingContainsNonFinite := E_Result.NotEvaluated;
        FExpectedContainsNaN := E_Result.Passed;
        FFindingContainsNaN := E_Result.NotEvaluated;
        FExpectedHasNoNaN := E_Result.Failed;
        FFindingHasNoNaN := E_Result.Failed;
        FExpectedContainsInfinity := E_Result.Failed;
        FFindingContainsInfinity := E_Result.Failed;
        FExpectedHasNoInfinity := E_Result.Passed;
        FFindingHasNoInfinity := E_Result.NotEvaluated;
    RowNaNLast:
        FValues[2] := FQuietNaN.Value;
        FExpectedIndex := 2;
        FExpectedAllElementsFinite := E_Result.Failed;
        FFindingAllElementsFinite := E_Result.Failed;
        FExpectedContainsNonFinite := E_Result.Passed;
        FFindingContainsNonFinite := E_Result.NotEvaluated;
        FExpectedContainsNaN := E_Result.Passed;
        FFindingContainsNaN := E_Result.NotEvaluated;
        FExpectedHasNoNaN := E_Result.Failed;
        FFindingHasNoNaN := E_Result.Failed;
        FExpectedContainsInfinity := E_Result.Failed;
        FFindingContainsInfinity := E_Result.Failed;
        FExpectedHasNoInfinity := E_Result.Passed;
        FFindingHasNoInfinity := E_Result.NotEvaluated;
    RowInfinityFirst:
        FValues[-2] := FPositiveInfinity.Value;
        FExpectedIndex := -2;
        FExpectedAllElementsFinite := E_Result.Failed;
        FFindingAllElementsFinite := E_Result.Failed;
        FExpectedContainsNonFinite := E_Result.Passed;
        FFindingContainsNonFinite := E_Result.NotEvaluated;
        FExpectedContainsNaN := E_Result.Failed;
        FFindingContainsNaN := E_Result.Failed;
        FExpectedHasNoNaN := E_Result.Passed;
        FFindingHasNoNaN := E_Result.NotEvaluated;
        FExpectedContainsInfinity := E_Result.Passed;
        FFindingContainsInfinity := E_Result.NotEvaluated;
        FExpectedHasNoInfinity := E_Result.Failed;
        FFindingHasNoInfinity := E_Result.Failed;
    RowInfinityMiddle:
        FValues[0] := FNegativeInfinity.Value;
        FExpectedIndex := 0;
        FExpectedAllElementsFinite := E_Result.Failed;
        FFindingAllElementsFinite := E_Result.Failed;
        FExpectedContainsNonFinite := E_Result.Passed;
        FFindingContainsNonFinite := E_Result.NotEvaluated;
        FExpectedContainsNaN := E_Result.Failed;
        FFindingContainsNaN := E_Result.Failed;
        FExpectedHasNoNaN := E_Result.Passed;
        FFindingHasNoNaN := E_Result.NotEvaluated;
        FExpectedContainsInfinity := E_Result.Passed;
        FFindingContainsInfinity := E_Result.NotEvaluated;
        FExpectedHasNoInfinity := E_Result.Failed;
        FFindingHasNoInfinity := E_Result.Failed;
    RowInfinityLast:
        FValues[2] := FPositiveInfinity.Value;
        FExpectedIndex := 2;
        FExpectedAllElementsFinite := E_Result.Failed;
        FFindingAllElementsFinite := E_Result.Failed;
        FExpectedContainsNonFinite := E_Result.Passed;
        FFindingContainsNonFinite := E_Result.NotEvaluated;
        FExpectedContainsNaN := E_Result.Failed;
        FFindingContainsNaN := E_Result.Failed;
        FExpectedHasNoNaN := E_Result.Passed;
        FFindingHasNoNaN := E_Result.NotEvaluated;
        FExpectedContainsInfinity := E_Result.Passed;
        FFindingContainsInfinity := E_Result.NotEvaluated;
        FExpectedHasNoInfinity := E_Result.Failed;
        FFindingHasNoInfinity := E_Result.Failed;
    RowMixedSpecials:
        FValues[-2] := FQuietNaN.Value;
        FValues[0] := FNegativeInfinity.Value;
        FExpectedIndex := -2;
        FExpectedInfinityIndex := 0;
        FExpectedAllElementsFinite := E_Result.Failed;
        FFindingAllElementsFinite := E_Result.Failed;
        FExpectedContainsNonFinite := E_Result.Passed;
        FFindingContainsNonFinite := E_Result.NotEvaluated;
        FExpectedContainsNaN := E_Result.Passed;
        FFindingContainsNaN := E_Result.NotEvaluated;
        FExpectedHasNoNaN := E_Result.Failed;
        FFindingHasNoNaN := E_Result.Failed;
        FExpectedContainsInfinity := E_Result.Passed;
        FFindingContainsInfinity := E_Result.NotEvaluated;
        FExpectedHasNoInfinity := E_Result.Failed;
        FFindingHasNoInfinity := E_Result.Failed;
    RowOutsideSelection:
        FValues[-2] := FQuietNaN.Value;
        FValues[2] := FPositiveInfinity.Value;
        FStartIndex := -1;
        FLength := 3;
        FExpectedAllElementsFinite := E_Result.Passed;
        FFindingAllElementsFinite := E_Result.NotEvaluated;
        FExpectedContainsNonFinite := E_Result.Failed;
        FFindingContainsNonFinite := E_Result.Failed;
        FExpectedContainsNaN := E_Result.Failed;
        FFindingContainsNaN := E_Result.Failed;
        FExpectedHasNoNaN := E_Result.Passed;
        FFindingHasNoNaN := E_Result.NotEvaluated;
        FExpectedContainsInfinity := E_Result.Failed;
        FFindingContainsInfinity := E_Result.Failed;
        FExpectedHasNoInfinity := E_Result.Passed;
        FFindingHasNoInfinity := E_Result.NotEvaluated;
    RowSingleLastElement:
        FValues[2] := FSignalingNaN.Value;
        FStartIndex := 2;
        FLength := 1;
        FExpectedIndex := 2;
        FExpectedAllElementsFinite := E_Result.Failed;
        FFindingAllElementsFinite := E_Result.Failed;
        FExpectedContainsNonFinite := E_Result.Passed;
        FFindingContainsNonFinite := E_Result.NotEvaluated;
        FExpectedContainsNaN := E_Result.Passed;
        FFindingContainsNaN := E_Result.NotEvaluated;
        FExpectedHasNoNaN := E_Result.Failed;
        FFindingHasNoNaN := E_Result.Failed;
        FExpectedContainsInfinity := E_Result.Failed;
        FFindingContainsInfinity := E_Result.Failed;
        FExpectedHasNoInfinity := E_Result.Passed;
        FFindingHasNoInfinity := E_Result.NotEvaluated;
    RowInvalidAfterFailed:
        FLength := 0;
        FPreserveResults := TRUE;
        FExpectedAllElementsFinite := E_Result.Error;
        FFindingAllElementsFinite := E_Result.Error;
        FExpectedContainsNonFinite := E_Result.Error;
        FFindingContainsNonFinite := E_Result.Error;
        FExpectedContainsNaN := E_Result.Error;
        FFindingContainsNaN := E_Result.Error;
        FExpectedHasNoNaN := E_Result.Error;
        FFindingHasNoNaN := E_Result.Error;
        FExpectedContainsInfinity := E_Result.Error;
        FFindingContainsInfinity := E_Result.Error;
        FExpectedHasNoInfinity := E_Result.Error;
        FFindingHasNoInfinity := E_Result.Error;
    RowErrorRemainsHeld:

        FPreserveResults := TRUE;
        FExpectedAllElementsFinite := E_Result.Error;
        FFindingAllElementsFinite := E_Result.NotEvaluated;
        FExpectedContainsNonFinite := E_Result.Error;
        FFindingContainsNonFinite := E_Result.NotEvaluated;
        FExpectedContainsNaN := E_Result.Error;
        FFindingContainsNaN := E_Result.NotEvaluated;
        FExpectedHasNoNaN := E_Result.Error;
        FFindingHasNoNaN := E_Result.NotEvaluated;
        FExpectedContainsInfinity := E_Result.Error;
        FFindingContainsInfinity := E_Result.NotEvaluated;
        FExpectedHasNoInfinity := E_Result.Error;
        FFindingHasNoInfinity := E_Result.NotEvaluated;
    RowStartBelowBounds:
        FStartIndex := -3;
        FExpectedAllElementsFinite := E_Result.Error;
        FFindingAllElementsFinite := E_Result.Error;
        FExpectedContainsNonFinite := E_Result.Error;
        FFindingContainsNonFinite := E_Result.Error;
        FExpectedContainsNaN := E_Result.Error;
        FFindingContainsNaN := E_Result.Error;
        FExpectedHasNoNaN := E_Result.Error;
        FFindingHasNoNaN := E_Result.Error;
        FExpectedContainsInfinity := E_Result.Error;
        FFindingContainsInfinity := E_Result.Error;
        FExpectedHasNoInfinity := E_Result.Error;
        FFindingHasNoInfinity := E_Result.Error;
    RowStartAboveBounds:
        FStartIndex := 3;
        FExpectedAllElementsFinite := E_Result.Error;
        FFindingAllElementsFinite := E_Result.Error;
        FExpectedContainsNonFinite := E_Result.Error;
        FFindingContainsNonFinite := E_Result.Error;
        FExpectedContainsNaN := E_Result.Error;
        FFindingContainsNaN := E_Result.Error;
        FExpectedHasNoNaN := E_Result.Error;
        FFindingHasNoNaN := E_Result.Error;
        FExpectedContainsInfinity := E_Result.Error;
        FFindingContainsInfinity := E_Result.Error;
        FExpectedHasNoInfinity := E_Result.Error;
        FFindingHasNoInfinity := E_Result.Error;
    RowEndAboveBounds:
        FStartIndex := 2;
        FLength := 2;
        FExpectedAllElementsFinite := E_Result.Error;
        FFindingAllElementsFinite := E_Result.Error;
        FExpectedContainsNonFinite := E_Result.Error;
        FFindingContainsNonFinite := E_Result.Error;
        FExpectedContainsNaN := E_Result.Error;
        FFindingContainsNaN := E_Result.Error;
        FExpectedHasNoNaN := E_Result.Error;
        FFindingHasNoNaN := E_Result.Error;
        FExpectedContainsInfinity := E_Result.Error;
        FFindingContainsInfinity := E_Result.Error;
        FExpectedHasNoInfinity := E_Result.Error;
        FFindingHasNoInfinity := E_Result.Error;
    RowLargeStart:
        FStartIndex := DINT#2147483647;
        FExpectedAllElementsFinite := E_Result.Error;
        FFindingAllElementsFinite := E_Result.Error;
        FExpectedContainsNonFinite := E_Result.Error;
        FFindingContainsNonFinite := E_Result.Error;
        FExpectedContainsNaN := E_Result.Error;
        FFindingContainsNaN := E_Result.Error;
        FExpectedHasNoNaN := E_Result.Error;
        FFindingHasNoNaN := E_Result.Error;
        FExpectedContainsInfinity := E_Result.Error;
        FFindingContainsInfinity := E_Result.Error;
        FExpectedHasNoInfinity := E_Result.Error;
        FFindingHasNoInfinity := E_Result.Error;
    RowZeroLength:
        FLength := 0;
        FExpectedAllElementsFinite := E_Result.Error;
        FFindingAllElementsFinite := E_Result.Error;
        FExpectedContainsNonFinite := E_Result.Error;
        FFindingContainsNonFinite := E_Result.Error;
        FExpectedContainsNaN := E_Result.Error;
        FFindingContainsNaN := E_Result.Error;
        FExpectedHasNoNaN := E_Result.Error;
        FFindingHasNoNaN := E_Result.Error;
        FExpectedContainsInfinity := E_Result.Error;
        FFindingContainsInfinity := E_Result.Error;
        FExpectedHasNoInfinity := E_Result.Error;
        FFindingHasNoInfinity := E_Result.Error;
    RowResetRecovers:

        FExpectedAllElementsFinite := E_Result.Passed;
        FFindingAllElementsFinite := E_Result.NotEvaluated;
        FExpectedContainsNonFinite := E_Result.Failed;
        FFindingContainsNonFinite := E_Result.Failed;
        FExpectedContainsNaN := E_Result.Failed;
        FFindingContainsNaN := E_Result.Failed;
        FExpectedHasNoNaN := E_Result.Passed;
        FFindingHasNoNaN := E_Result.NotEvaluated;
        FExpectedContainsInfinity := E_Result.Failed;
        FFindingContainsInfinity := E_Result.Failed;
        FExpectedHasNoInfinity := E_Result.Passed;
        FFindingHasNoInfinity := E_Result.NotEvaluated;
ELSE
    Error(Message := 'Unknown classification selftest row.');
END_CASE;
END_METHOD

END_FUNCTION_BLOCK

// ---- Framework/Assertions/POU/Arrays/LReal/AssertArrayAllElementsFinite_LReal.TcPOU
{region 'Documentation'}
(*!
<summary>Checks that every selected element is finite.</summary>
<description>

Invalid binding/range is Error; a classification mismatch is Failed. Only the selected
range is inspected.

StartIndex is an absolute declared IN index, not an offset. Length selects 1..255
elements; the complete selected range must fit IN. Invalid references or ranges report
Error.

Keep supplied arrays stable for the call. Input data is read, not copied or retained as a
snapshot.

NaN and either infinity are legitimate checked data, not configuration errors.
Classification mismatch reports Failed. Bit-based classification does not perform an ordered
floating-point comparison.

Numeric diagnostics use the formatter's default six significant digits; rounding affects
the message only, not the comparison.

</description>
*)
{endregion}
FUNCTION_BLOCK AssertArrayAllElementsFinite_LReal EXTENDS AssertionBase
VAR_INPUT
    StartIndex : DINT; //! First selected index in IN; uses the array's declared index range, not a zero-based offset.
    Length : USINT; //! Number of inspected elements, from 1 through 255.
END_VAR
VAR_IN_OUT CONSTANT
    IN : ARRAY[*] OF LREAL; //! Read-only checked data; keep stable during the call.
END_VAR

SUPER^();

{region 'Documentation'}
(*!
<summary>Validates the selected range, then classifies element representations.</summary>
*)
{endregion}
METHOD PROTECTED Assert
VAR
    InLowerIndex : DINT;
    InUpperIndex : DINT;
    EndIndex : LINT;
    Offset : LINT;
    InIndex : DINT;
    ValueFound : BOOL;
    Representation : AssertionLRealRepresentation;
    Message : STRING(GVL_Constants.MessageLength);
END_VAR
VAR CONSTANT
    ExponentMask : LWORD := LWORD#16#7FF0000000000000;
END_VAR
IF NOT EvaluationActive THEN
    RETURN;
END_IF;

IF Result = E_Result.Error THEN
    RETURN;
END_IF;

// C0371: FB input is checked here before any reference access.
{warning disable C0371}
IF NOT __ISVALIDREF(IN) THEN
    Error(Message := 'Assertion error: IN reference is invalid.');
    RETURN;
END_IF;

InLowerIndex := LOWER_BOUND(IN, 1);
InUpperIndex := UPPER_BOUND(IN, 1);
EndIndex := DINT_TO_LINT(StartIndex) + USINT_TO_LINT(Length) - 1;

IF (Length = 0)
    OR (StartIndex < InLowerIndex) OR (StartIndex > InUpperIndex)
    OR (EndIndex > DINT_TO_LINT(InUpperIndex)) THEN
    Message := CONCAT('Assertion error: array range is invalid. StartIndex = ',
        DINT_TO_STRING(StartIndex));
    Message := CONCAT(Message, ', Length = ');
    Message := CONCAT(Message, USINT_TO_STRING(Length));
    Message := CONCAT(Message, '.');
    Error(Message := Message);
    RETURN;
END_IF;

IF Result = E_Result.Failed THEN
    RETURN;
END_IF;

ValueFound := FALSE;
FOR Offset := 0 TO USINT_TO_LINT(Length) - 1 DO
    InIndex := LINT_TO_DINT(DINT_TO_LINT(StartIndex) + Offset);
    Representation.Value := IN[InIndex];
    ValueFound := (Representation.Bits AND ExponentMask) = ExponentMask;
    IF ValueFound THEN
        EXIT;
    END_IF;
END_FOR;

IF ValueFound THEN
    Message := 'Assertion failed: array range contains a non-finite value.';
    Message := CONCAT(Message, ' Actual[');
    Message := CONCAT(Message, DINT_TO_STRING(InIndex));
    Message := CONCAT(Message, '] = ');
    Message := CONCAT(Message, CreateAssertionTextValue_LReal(Value := Representation.Value));
    Message := CONCAT(Message, ', Range = [');
    Message := CONCAT(Message, DINT_TO_STRING(StartIndex));
    Message := CONCAT(Message, '..');
    Message := CONCAT(Message, LINT_TO_STRING(EndIndex));
    Message := CONCAT(Message, '].');
    Fail(Message := Message);
    RETURN;
END_IF;

Pass();
{warning restore C0371}
END_METHOD

END_FUNCTION_BLOCK

// ---- Framework/Assertions/POU/Arrays/LReal/AssertArrayContainsNonFinite_LReal.TcPOU
{region 'Documentation'}
(*!
<summary>Checks that the selected range contains NaN or either infinity.</summary>
<description>

Invalid binding/range is Error; a classification mismatch is Failed. Only the selected
range is inspected.

StartIndex is an absolute declared IN index, not an offset. Length selects 1..255
elements; the complete selected range must fit IN. Invalid references or ranges report
Error.

Keep supplied arrays stable for the call. Input data is read, not copied or retained as a
snapshot.

NaN and either infinity are legitimate checked data, not configuration errors.
Classification mismatch reports Failed. Bit-based classification does not perform an ordered
floating-point comparison.

</description>
*)
{endregion}
FUNCTION_BLOCK AssertArrayContainsNonFinite_LReal EXTENDS AssertionBase
VAR_INPUT
    StartIndex : DINT; //! First selected index in IN; uses the array's declared index range, not a zero-based offset.
    Length : USINT; //! Number of inspected elements, from 1 through 255.
END_VAR
VAR_IN_OUT CONSTANT
    IN : ARRAY[*] OF LREAL; //! Read-only checked data; keep stable during the call.
END_VAR

SUPER^();

{region 'Documentation'}
(*!
<summary>Validates the selected range, then classifies element representations.</summary>
*)
{endregion}
METHOD PROTECTED Assert
VAR
    InLowerIndex : DINT;
    InUpperIndex : DINT;
    EndIndex : LINT;
    Offset : LINT;
    InIndex : DINT;
    ValueFound : BOOL;
    Representation : AssertionLRealRepresentation;
    Message : STRING(GVL_Constants.MessageLength);
END_VAR
VAR CONSTANT
    ExponentMask : LWORD := LWORD#16#7FF0000000000000;
END_VAR
IF NOT EvaluationActive THEN
    RETURN;
END_IF;

IF Result = E_Result.Error THEN
    RETURN;
END_IF;

// C0371: FB input is checked here before any reference access.
{warning disable C0371}
IF NOT __ISVALIDREF(IN) THEN
    Error(Message := 'Assertion error: IN reference is invalid.');
    RETURN;
END_IF;

InLowerIndex := LOWER_BOUND(IN, 1);
InUpperIndex := UPPER_BOUND(IN, 1);
EndIndex := DINT_TO_LINT(StartIndex) + USINT_TO_LINT(Length) - 1;

IF (Length = 0)
    OR (StartIndex < InLowerIndex) OR (StartIndex > InUpperIndex)
    OR (EndIndex > DINT_TO_LINT(InUpperIndex)) THEN
    Message := CONCAT('Assertion error: array range is invalid. StartIndex = ',
        DINT_TO_STRING(StartIndex));
    Message := CONCAT(Message, ', Length = ');
    Message := CONCAT(Message, USINT_TO_STRING(Length));
    Message := CONCAT(Message, '.');
    Error(Message := Message);
    RETURN;
END_IF;

IF Result = E_Result.Failed THEN
    RETURN;
END_IF;

ValueFound := FALSE;
FOR Offset := 0 TO USINT_TO_LINT(Length) - 1 DO
    InIndex := LINT_TO_DINT(DINT_TO_LINT(StartIndex) + Offset);
    Representation.Value := IN[InIndex];
    ValueFound := (Representation.Bits AND ExponentMask) = ExponentMask;
    IF ValueFound THEN
        EXIT;
    END_IF;
END_FOR;

IF NOT ValueFound THEN
    Message := 'Assertion failed: array range contains no non-finite value.';
    Message := CONCAT(Message, ', Range = [');
    Message := CONCAT(Message, DINT_TO_STRING(StartIndex));
    Message := CONCAT(Message, '..');
    Message := CONCAT(Message, LINT_TO_STRING(EndIndex));
    Message := CONCAT(Message, '].');
    Fail(Message := Message);
    RETURN;
END_IF;

Pass();
{warning restore C0371}
END_METHOD

END_FUNCTION_BLOCK

// ---- Framework/Assertions/POU/Arrays/LReal/AssertArrayContainsNaN_LReal.TcPOU
{region 'Documentation'}
(*!
<summary>Checks that the selected range contains NaN.</summary>
<description>

Invalid binding/range is Error; a classification mismatch is Failed. Only the selected
range is inspected.

StartIndex is an absolute declared IN index, not an offset. Length selects 1..255
elements; the complete selected range must fit IN. Invalid references or ranges report
Error.

Keep supplied arrays stable for the call. Input data is read, not copied or retained as a
snapshot.

NaN and either infinity are legitimate checked data, not configuration errors.
Classification mismatch reports Failed. Bit-based classification does not perform an ordered
floating-point comparison.

</description>
*)
{endregion}
FUNCTION_BLOCK AssertArrayContainsNaN_LReal EXTENDS AssertionBase
VAR_INPUT
    StartIndex : DINT; //! First selected index in IN; uses the array's declared index range, not a zero-based offset.
    Length : USINT; //! Number of inspected elements, from 1 through 255.
END_VAR
VAR_IN_OUT CONSTANT
    IN : ARRAY[*] OF LREAL; //! Read-only checked data; keep stable during the call.
END_VAR

SUPER^();

{region 'Documentation'}
(*!
<summary>Validates the selected range, then classifies element representations.</summary>
*)
{endregion}
METHOD PROTECTED Assert
VAR
    InLowerIndex : DINT;
    InUpperIndex : DINT;
    EndIndex : LINT;
    Offset : LINT;
    InIndex : DINT;
    ValueFound : BOOL;
    Representation : AssertionLRealRepresentation;
    Message : STRING(GVL_Constants.MessageLength);
END_VAR
VAR CONSTANT
    ExponentMask : LWORD := LWORD#16#7FF0000000000000;
    FractionMask : LWORD := LWORD#16#000FFFFFFFFFFFFF;
END_VAR
IF NOT EvaluationActive THEN
    RETURN;
END_IF;

IF Result = E_Result.Error THEN
    RETURN;
END_IF;

// C0371: FB input is checked here before any reference access.
{warning disable C0371}
IF NOT __ISVALIDREF(IN) THEN
    Error(Message := 'Assertion error: IN reference is invalid.');
    RETURN;
END_IF;

InLowerIndex := LOWER_BOUND(IN, 1);
InUpperIndex := UPPER_BOUND(IN, 1);
EndIndex := DINT_TO_LINT(StartIndex) + USINT_TO_LINT(Length) - 1;

IF (Length = 0)
    OR (StartIndex < InLowerIndex) OR (StartIndex > InUpperIndex)
    OR (EndIndex > DINT_TO_LINT(InUpperIndex)) THEN
    Message := CONCAT('Assertion error: array range is invalid. StartIndex = ',
        DINT_TO_STRING(StartIndex));
    Message := CONCAT(Message, ', Length = ');
    Message := CONCAT(Message, USINT_TO_STRING(Length));
    Message := CONCAT(Message, '.');
    Error(Message := Message);
    RETURN;
END_IF;

IF Result = E_Result.Failed THEN
    RETURN;
END_IF;

ValueFound := FALSE;
FOR Offset := 0 TO USINT_TO_LINT(Length) - 1 DO
    InIndex := LINT_TO_DINT(DINT_TO_LINT(StartIndex) + Offset);
    Representation.Value := IN[InIndex];
    ValueFound := ((Representation.Bits AND ExponentMask) = ExponentMask)
        AND ((Representation.Bits AND FractionMask) <> 0);
    IF ValueFound THEN
        EXIT;
    END_IF;
END_FOR;

IF NOT ValueFound THEN
    Message := 'Assertion failed: array range contains no NaN.';
    Message := CONCAT(Message, ', Range = [');
    Message := CONCAT(Message, DINT_TO_STRING(StartIndex));
    Message := CONCAT(Message, '..');
    Message := CONCAT(Message, LINT_TO_STRING(EndIndex));
    Message := CONCAT(Message, '].');
    Fail(Message := Message);
    RETURN;
END_IF;

Pass();
{warning restore C0371}
END_METHOD

END_FUNCTION_BLOCK

// ---- Framework/Assertions/POU/Arrays/LReal/AssertArrayHasNoNaN_LReal.TcPOU
{region 'Documentation'}
(*!
<summary>Checks that the selected range contains no NaN; infinities are allowed.</summary>
<description>

Invalid binding/range is Error; a classification mismatch is Failed. Only the selected
range is inspected.

StartIndex is an absolute declared IN index, not an offset. Length selects 1..255
elements; the complete selected range must fit IN. Invalid references or ranges report
Error.

Keep supplied arrays stable for the call. Input data is read, not copied or retained as a
snapshot.

NaN and either infinity are legitimate checked data, not configuration errors.
Classification mismatch reports Failed. Bit-based classification does not perform an ordered
floating-point comparison.

Numeric diagnostics use the formatter's default six significant digits; rounding affects
the message only, not the comparison.

</description>
*)
{endregion}
FUNCTION_BLOCK AssertArrayHasNoNaN_LReal EXTENDS AssertionBase
VAR_INPUT
    StartIndex : DINT; //! First selected index in IN; uses the array's declared index range, not a zero-based offset.
    Length : USINT; //! Number of inspected elements, from 1 through 255.
END_VAR
VAR_IN_OUT CONSTANT
    IN : ARRAY[*] OF LREAL; //! Read-only checked data; keep stable during the call.
END_VAR

SUPER^();

{region 'Documentation'}
(*!
<summary>Validates the selected range, then classifies element representations.</summary>
*)
{endregion}
METHOD PROTECTED Assert
VAR
    InLowerIndex : DINT;
    InUpperIndex : DINT;
    EndIndex : LINT;
    Offset : LINT;
    InIndex : DINT;
    ValueFound : BOOL;
    Representation : AssertionLRealRepresentation;
    Message : STRING(GVL_Constants.MessageLength);
END_VAR
VAR CONSTANT
    ExponentMask : LWORD := LWORD#16#7FF0000000000000;
    FractionMask : LWORD := LWORD#16#000FFFFFFFFFFFFF;
END_VAR
IF NOT EvaluationActive THEN
    RETURN;
END_IF;

IF Result = E_Result.Error THEN
    RETURN;
END_IF;

// C0371: FB input is checked here before any reference access.
{warning disable C0371}
IF NOT __ISVALIDREF(IN) THEN
    Error(Message := 'Assertion error: IN reference is invalid.');
    RETURN;
END_IF;

InLowerIndex := LOWER_BOUND(IN, 1);
InUpperIndex := UPPER_BOUND(IN, 1);
EndIndex := DINT_TO_LINT(StartIndex) + USINT_TO_LINT(Length) - 1;

IF (Length = 0)
    OR (StartIndex < InLowerIndex) OR (StartIndex > InUpperIndex)
    OR (EndIndex > DINT_TO_LINT(InUpperIndex)) THEN
    Message := CONCAT('Assertion error: array range is invalid. StartIndex = ',
        DINT_TO_STRING(StartIndex));
    Message := CONCAT(Message, ', Length = ');
    Message := CONCAT(Message, USINT_TO_STRING(Length));
    Message := CONCAT(Message, '.');
    Error(Message := Message);
    RETURN;
END_IF;

IF Result = E_Result.Failed THEN
    RETURN;
END_IF;

ValueFound := FALSE;
FOR Offset := 0 TO USINT_TO_LINT(Length) - 1 DO
    InIndex := LINT_TO_DINT(DINT_TO_LINT(StartIndex) + Offset);
    Representation.Value := IN[InIndex];
    ValueFound := ((Representation.Bits AND ExponentMask) = ExponentMask)
        AND ((Representation.Bits AND FractionMask) <> 0);
    IF ValueFound THEN
        EXIT;
    END_IF;
END_FOR;

IF ValueFound THEN
    Message := 'Assertion failed: array range contains NaN.';
    Message := CONCAT(Message, ' Actual[');
    Message := CONCAT(Message, DINT_TO_STRING(InIndex));
    Message := CONCAT(Message, '] = ');
    Message := CONCAT(Message, CreateAssertionTextValue_LReal(Value := Representation.Value));
    Message := CONCAT(Message, ', Range = [');
    Message := CONCAT(Message, DINT_TO_STRING(StartIndex));
    Message := CONCAT(Message, '..');
    Message := CONCAT(Message, LINT_TO_STRING(EndIndex));
    Message := CONCAT(Message, '].');
    Fail(Message := Message);
    RETURN;
END_IF;

Pass();
{warning restore C0371}
END_METHOD

END_FUNCTION_BLOCK

// ---- Framework/Assertions/POU/Arrays/LReal/AssertArrayContainsInfinity_LReal.TcPOU
{region 'Documentation'}
(*!
<summary>Checks that the selected range contains either infinity.</summary>
<description>

Invalid binding/range is Error; a classification mismatch is Failed. Only the selected
range is inspected.

StartIndex is an absolute declared IN index, not an offset. Length selects 1..255
elements; the complete selected range must fit IN. Invalid references or ranges report
Error.

Keep supplied arrays stable for the call. Input data is read, not copied or retained as a
snapshot.

NaN and either infinity are legitimate checked data, not configuration errors.
Classification mismatch reports Failed. Bit-based classification does not perform an ordered
floating-point comparison.

</description>
*)
{endregion}
FUNCTION_BLOCK AssertArrayContainsInfinity_LReal EXTENDS AssertionBase
VAR_INPUT
    StartIndex : DINT; //! First selected index in IN; uses the array's declared index range, not a zero-based offset.
    Length : USINT; //! Number of inspected elements, from 1 through 255.
END_VAR
VAR_IN_OUT CONSTANT
    IN : ARRAY[*] OF LREAL; //! Read-only checked data; keep stable during the call.
END_VAR

SUPER^();

{region 'Documentation'}
(*!
<summary>Validates the selected range, then classifies element representations.</summary>
*)
{endregion}
METHOD PROTECTED Assert
VAR
    InLowerIndex : DINT;
    InUpperIndex : DINT;
    EndIndex : LINT;
    Offset : LINT;
    InIndex : DINT;
    ValueFound : BOOL;
    Representation : AssertionLRealRepresentation;
    Message : STRING(GVL_Constants.MessageLength);
END_VAR
VAR CONSTANT
    ExponentMask : LWORD := LWORD#16#7FF0000000000000;
    FractionMask : LWORD := LWORD#16#000FFFFFFFFFFFFF;
END_VAR
IF NOT EvaluationActive THEN
    RETURN;
END_IF;

IF Result = E_Result.Error THEN
    RETURN;
END_IF;

// C0371: FB input is checked here before any reference access.
{warning disable C0371}
IF NOT __ISVALIDREF(IN) THEN
    Error(Message := 'Assertion error: IN reference is invalid.');
    RETURN;
END_IF;

InLowerIndex := LOWER_BOUND(IN, 1);
InUpperIndex := UPPER_BOUND(IN, 1);
EndIndex := DINT_TO_LINT(StartIndex) + USINT_TO_LINT(Length) - 1;

IF (Length = 0)
    OR (StartIndex < InLowerIndex) OR (StartIndex > InUpperIndex)
    OR (EndIndex > DINT_TO_LINT(InUpperIndex)) THEN
    Message := CONCAT('Assertion error: array range is invalid. StartIndex = ',
        DINT_TO_STRING(StartIndex));
    Message := CONCAT(Message, ', Length = ');
    Message := CONCAT(Message, USINT_TO_STRING(Length));
    Message := CONCAT(Message, '.');
    Error(Message := Message);
    RETURN;
END_IF;

IF Result = E_Result.Failed THEN
    RETURN;
END_IF;

ValueFound := FALSE;
FOR Offset := 0 TO USINT_TO_LINT(Length) - 1 DO
    InIndex := LINT_TO_DINT(DINT_TO_LINT(StartIndex) + Offset);
    Representation.Value := IN[InIndex];
    ValueFound := ((Representation.Bits AND ExponentMask) = ExponentMask)
        AND ((Representation.Bits AND FractionMask) = 0);
    IF ValueFound THEN
        EXIT;
    END_IF;
END_FOR;

IF NOT ValueFound THEN
    Message := 'Assertion failed: array range contains no infinity.';
    Message := CONCAT(Message, ', Range = [');
    Message := CONCAT(Message, DINT_TO_STRING(StartIndex));
    Message := CONCAT(Message, '..');
    Message := CONCAT(Message, LINT_TO_STRING(EndIndex));
    Message := CONCAT(Message, '].');
    Fail(Message := Message);
    RETURN;
END_IF;

Pass();
{warning restore C0371}
END_METHOD

END_FUNCTION_BLOCK

// ---- Framework/Assertions/POU/Arrays/LReal/AssertArrayHasNoInfinity_LReal.TcPOU
{region 'Documentation'}
(*!
<summary>Checks that the selected range contains no infinity; NaN is allowed.</summary>
<description>

Invalid binding/range is Error; a classification mismatch is Failed. Only the selected
range is inspected.

StartIndex is an absolute declared IN index, not an offset. Length selects 1..255
elements; the complete selected range must fit IN. Invalid references or ranges report
Error.

Keep supplied arrays stable for the call. Input data is read, not copied or retained as a
snapshot.

NaN and either infinity are legitimate checked data, not configuration errors.
Classification mismatch reports Failed. Bit-based classification does not perform an ordered
floating-point comparison.

Numeric diagnostics use the formatter's default six significant digits; rounding affects
the message only, not the comparison.

</description>
*)
{endregion}
FUNCTION_BLOCK AssertArrayHasNoInfinity_LReal EXTENDS AssertionBase
VAR_INPUT
    StartIndex : DINT; //! First selected index in IN; uses the array's declared index range, not a zero-based offset.
    Length : USINT; //! Number of inspected elements, from 1 through 255.
END_VAR
VAR_IN_OUT CONSTANT
    IN : ARRAY[*] OF LREAL; //! Read-only checked data; keep stable during the call.
END_VAR

SUPER^();

{region 'Documentation'}
(*!
<summary>Validates the selected range, then classifies element representations.</summary>
*)
{endregion}
METHOD PROTECTED Assert
VAR
    InLowerIndex : DINT;
    InUpperIndex : DINT;
    EndIndex : LINT;
    Offset : LINT;
    InIndex : DINT;
    ValueFound : BOOL;
    Representation : AssertionLRealRepresentation;
    Message : STRING(GVL_Constants.MessageLength);
END_VAR
VAR CONSTANT
    ExponentMask : LWORD := LWORD#16#7FF0000000000000;
    FractionMask : LWORD := LWORD#16#000FFFFFFFFFFFFF;
END_VAR
IF NOT EvaluationActive THEN
    RETURN;
END_IF;

IF Result = E_Result.Error THEN
    RETURN;
END_IF;

// C0371: FB input is checked here before any reference access.
{warning disable C0371}
IF NOT __ISVALIDREF(IN) THEN
    Error(Message := 'Assertion error: IN reference is invalid.');
    RETURN;
END_IF;

InLowerIndex := LOWER_BOUND(IN, 1);
InUpperIndex := UPPER_BOUND(IN, 1);
EndIndex := DINT_TO_LINT(StartIndex) + USINT_TO_LINT(Length) - 1;

IF (Length = 0)
    OR (StartIndex < InLowerIndex) OR (StartIndex > InUpperIndex)
    OR (EndIndex > DINT_TO_LINT(InUpperIndex)) THEN
    Message := CONCAT('Assertion error: array range is invalid. StartIndex = ',
        DINT_TO_STRING(StartIndex));
    Message := CONCAT(Message, ', Length = ');
    Message := CONCAT(Message, USINT_TO_STRING(Length));
    Message := CONCAT(Message, '.');
    Error(Message := Message);
    RETURN;
END_IF;

IF Result = E_Result.Failed THEN
    RETURN;
END_IF;

ValueFound := FALSE;
FOR Offset := 0 TO USINT_TO_LINT(Length) - 1 DO
    InIndex := LINT_TO_DINT(DINT_TO_LINT(StartIndex) + Offset);
    Representation.Value := IN[InIndex];
    ValueFound := ((Representation.Bits AND ExponentMask) = ExponentMask)
        AND ((Representation.Bits AND FractionMask) = 0);
    IF ValueFound THEN
        EXIT;
    END_IF;
END_FOR;

IF ValueFound THEN
    Message := 'Assertion failed: array range contains infinity.';
    Message := CONCAT(Message, ' Actual[');
    Message := CONCAT(Message, DINT_TO_STRING(InIndex));
    Message := CONCAT(Message, '] = ');
    Message := CONCAT(Message, CreateAssertionTextValue_LReal(Value := Representation.Value));
    Message := CONCAT(Message, ', Range = [');
    Message := CONCAT(Message, DINT_TO_STRING(StartIndex));
    Message := CONCAT(Message, '..');
    Message := CONCAT(Message, LINT_TO_STRING(EndIndex));
    Message := CONCAT(Message, '].');
    Fail(Message := Message);
    RETURN;
END_IF;

Pass();
{warning restore C0371}
END_METHOD

END_FUNCTION_BLOCK

// ---- SelfTests/TestSuites/TestSuite_AssertionObservation.TcPOU
{region 'Documentation'}
(*!
<summary>Checks temporal Assertion observation with isolated, deterministic cycle traces.</summary>
*)
{endregion}
FUNCTION_BLOCK TestSuite_AssertionObservation EXTENDS TestSuiteBase
VAR
    FEdgeObservation : Test_AssertionEdgeObservation;
    FEdgeCount : Test_AssertionEdgeCount;
    FSequence : Test_AssertionSequence;
    FScalarObservation : Test_AssertionScalarObservation;
    FArraySnapshot : Test_AssertionArraySnapshot;
    FFloatingSnapshot : Test_AssertionFloatingSnapshot;
    FTestCases : ARRAY[1..TestCaseCapacity] OF I_TestCase;
END_VAR
VAR CONSTANT
    TestCaseCapacity : UINT := 6;
END_VAR

SUPER^();

{region 'Documentation'}
(*!
<summary>Initializes six isolated observation scenarios and registers them serially.</summary>
*)
{endregion}
METHOD PROTECTED Configure
VAR_IN_OUT
    // SA0167: Borrowed owner builder; no temporary instance is created.
    {attribute 'analysis' := '-167'}
    Builder : TestSuiteConfigurationBuilder; //! Borrowed owner configuration builder used only during this Configure call; register this owner's concrete children.
END_VAR
VAR
    TestConfig : ST_TestCaseConfig;
END_VAR
Builder.Initialize(Mode := E_OrchestrationMode.Serial,
    TestCases := FTestCases);
FEdgeObservation.Initialize(Parent := THIS^,
    TestName := 'EdgeObservation',
    Config := TestConfig);
Builder.Register(TestCase := FEdgeObservation);
FEdgeCount.Initialize(Parent := THIS^,
    TestName := 'EdgeCount',
    Config := TestConfig);
Builder.Register(TestCase := FEdgeCount);
FSequence.Initialize(Parent := THIS^,
    TestName := 'Sequence',
    Config := TestConfig);
Builder.Register(TestCase := FSequence);
FScalarObservation.Initialize(Parent := THIS^,
    TestName := 'ScalarObservation',
    Config := TestConfig);
Builder.Register(TestCase := FScalarObservation);
FArraySnapshot.Initialize(Parent := THIS^,
    TestName := 'ArraySnapshot',
    Config := TestConfig);
Builder.Register(TestCase := FArraySnapshot);
FFloatingSnapshot.Initialize(Parent := THIS^,
    TestName := 'FloatingSnapshot',
    Config := TestConfig);
Builder.Register(TestCase := FFloatingSnapshot);
END_METHOD

{region 'Documentation'}
(*!
<summary>Returns a registered scenario using its original array index.</summary>
*)
{endregion}
METHOD PUBLIC GetTestCase : I_TestCase //! Typed child interface at the original array index; zero when no entry is available.
VAR_INPUT
    Index : DINT; //! Original occupied child-array index, rather than an ordinal position.
END_VAR
GetTestCase := 0;
IF (ChildCount = 0) OR (Index < ChildArrayLowerBound)
    OR (DINT_TO_LINT(Index) >= DINT_TO_LINT(ChildArrayLowerBound) + UINT_TO_LINT(ChildCount)) THEN
    RETURN;
END_IF;
GetTestCase := FTestCases[Index];
END_METHOD

{region 'Documentation'}
(*!
<summary>Calls every owned scenario once per initialized Suite cycle.</summary>
*)
{endregion}
METHOD PROTECTED ProcessTestCases
FEdgeObservation();
FEdgeCount();
FSequence();
FScalarObservation();
FArraySnapshot();
FFloatingSnapshot();
END_METHOD

END_FUNCTION_BLOCK

// ---- SelfTests/TestCases/TestSuite_AssertionObservation/Test_AssertionEdgeObservation.TcPOU
{region 'Documentation'}
(*!
<summary>Checks rising/falling edge baselines, interruptions and delayed observation.</summary>
<description>
Normal and delayed subjects receive mirrored signals so both edge directions have the same literal expectations. A disabled call breaks sample adjacency; the held result survives. Delayed subjects use ObserveFirstCycle FALSE. No adapter overrides production observation logic.
ProcessTests executes one named step per PLC cycle. ProcessAssertions checks that
step before the next call advances it. Every trace has its own outer Assertion;
FirstFailedStep retains the first mismatching checkpoint for online diagnosis.
Expected findings are captured locally and checked before the next step clears
that capture. Subjects are deliberately not called between scripted steps.
</description>
*)
{endregion}
FUNCTION_BLOCK Test_AssertionEdgeObservation EXTENDS TestCaseBase
VAR
    FRising : AssertNoRisingEdge;
    FFalling : AssertNoFallingEdge;
    FDelayedRising : AssertNoRisingEdge;
    FDelayedFalling : AssertNoFallingEdge;
    FCapture : EventBuffer;
    FEvents : ARRAY[1..CaptureLength] OF ST_Event;
    FCaptureFifo : ST_FifoStatus;
    FCaptureStatus : ST_EventBufferStatus;
    FSetupValid : BOOL;
    FStep : UINT;
    FTrace : UINT;
    FFirstFailedStep : UINT;
    FChecked : BOOL;
    FObservationReady : BOOL;
    FStepMatches : BOOL;
    FResultsMatch : BOOL;
    FActivityMatches : BOOL;
    FFindingsMatch : BOOL;
    FSample : BOOL;
    FSubjectEnable : BOOL;
    FResetSubjects : BOOL;
    FExpectedResult : E_Result;
    FExpectedDelayedResult : E_Result;
    FExpectedObservation : BOOL;
    FExpectedDelayedObservation : BOOL;
    FExpectedEvaluation : BOOL;
    FExpectedDelayedEvaluation : BOOL;
    FRisingFindingExpected : BOOL;
    FFallingFindingExpected : BOOL;
    FDelayedRisingFindingExpected : BOOL;
    FDelayedFallingFindingExpected : BOOL;
END_VAR
VAR
    FResetHistory : AssertTrue;
    FFirstObservation : AssertTrue;
    FHeldFailure : AssertTrue;
    FDisabledHistory : AssertTrue;
    FDelayedObservation : AssertTrue;
END_VAR
VAR CONSTANT
    CaptureLength : UINT := 8;
    StepInitialBoundReset : UINT := 1;
    StepFirstHighSample : UINT := 2;
    StepSameHighSample : UINT := 3;
    StepOppositeEdgeAllowed : UINT := 4;
    StepForbiddenEdge : UINT := 5;
    StepRepeatedFailure : UINT := 6;
    StepResetBeforeGap : UINT := 7;
    StepBaselineBeforeGap : UINT := 8;
    StepDisabledChange : UINT := 9;
    StepFirstAfterGap : UINT := 10;
    StepSecondAfterGap : UINT := 11;
    StepAllowedAfterGap : UINT := 12;
    StepForbiddenAfterGap : UINT := 13;
    StepResetBeforeDelay : UINT := 14;
    StepSkippedFirstBaseline : UINT := 15;
    StepEdgeBeforeDelayedBaseline : UINT := 16;
    StepStableDelayedBaseline : UINT := 17;
    LastStep : UINT := StepStableDelayedBaseline;
    TraceResetHistory : UINT := 1;
    TraceFirstObservation : UINT := 2;
    TraceHeldFailure : UINT := 3;
    TraceDisabledHistory : UINT := 4;
    TraceDelayedObservation : UINT := 5;
END_VAR

SUPER^();

{region 'Documentation'}
(*!
<summary>Collects the outer trace checks, never subject results.</summary>
*)
{endregion}
METHOD PROTECTED AggregateResults
VAR_INPUT
    Aggregator : I_ResultAggregator; //! Borrowed result sink owned by the outer Test Case; add this test's checking Assertions without resetting or retaining the sink.
END_VAR
Aggregator.AddProvider(Provider := FResetHistory);
Aggregator.AddProvider(Provider := FFirstObservation);
Aggregator.AddProvider(Provider := FHeldFailure);
Aggregator.AddProvider(Provider := FDisabledHistory);
Aggregator.AddProvider(Provider := FDelayedObservation);
END_METHOD

{region 'Documentation'}
(*!
<summary>Calls each real production subject once with this step's bound inputs.</summary>
*)
{endregion}
METHOD PRIVATE CallSubjects
FRising(Enable := FSubjectEnable,
    State := E_State.Running,
    IN := FSample);
FFalling(Enable := FSubjectEnable,
    State := E_State.Running,
    IN := NOT FSample);
FDelayedRising(Enable := FSubjectEnable,
    State := E_State.Running,
    IN := FSample);
FDelayedFalling(Enable := FSubjectEnable,
    State := E_State.Running,
    IN := NOT FSample);
END_METHOD

{region 'Documentation'}
(*!
<summary>Checks per-step finding order, identity and count without retaining old events.</summary>
*)
{endregion}
METHOD PRIVATE CheckFindings
VAR
    Index : UINT;
    FindingMatches : BOOL;
END_VAR
Index := 1;
FFindingsMatch := TRUE;
IF FRisingFindingExpected THEN
    FindingMatches := IsFindingValid(Index := Index,
        ExpectedName := FRising.Name);
    FFindingsMatch := FFindingsMatch AND FindingMatches;
    Index := Index + 1;
END_IF;
IF FFallingFindingExpected THEN
    FindingMatches := IsFindingValid(Index := Index,
        ExpectedName := FFalling.Name);
    FFindingsMatch := FFindingsMatch AND FindingMatches;
    Index := Index + 1;
END_IF;
IF FDelayedRisingFindingExpected THEN
    FindingMatches := IsFindingValid(Index := Index,
        ExpectedName := FDelayedRising.Name);
    FFindingsMatch := FFindingsMatch AND FindingMatches;
    Index := Index + 1;
END_IF;
IF FDelayedFallingFindingExpected THEN
    FindingMatches := IsFindingValid(Index := Index,
        ExpectedName := FDelayedFalling.Name);
    FFindingsMatch := FFindingsMatch AND FindingMatches;
    Index := Index + 1;
END_IF;
FFindingsMatch := FFindingsMatch
    AND (FCaptureStatus.SequenceId = UINT_TO_UDINT(Index - 1))
    AND (FCaptureStatus.LostEventCount = 0);
END_METHOD

{region 'Documentation'}
(*!
<summary>Rejects incomplete local capture, subject or checking-Assertion setup.</summary>
*)
{endregion}
METHOD PROTECTED CheckInitialization : BOOL //! TRUE when the inherited initialization check and this concrete fixture check both accept the setup.
CheckInitialization := SUPER^.CheckInitialization();
IF NOT CheckInitialization THEN
    RETURN;
END_IF;

CheckInitialization := FSetupValid
    AND FResetHistory.IsInitialized
    AND FFirstObservation.IsInitialized
    AND FHeldFailure.IsInitialized
    AND FDisabledHistory.IsInitialized
    AND FDelayedObservation.IsInitialized;
IF NOT CheckInitialization THEN
    EventPublisher.PublishEvent(Event := CreateFrameworkEvent(Name := Name,
        ResourceName := '',
        State := State,
        Severity := E_EventSeverity.Error,
        Message := 'Observation selftest setup failed.'));
END_IF;
END_METHOD

{region 'Documentation'}
(*!
<summary>Compares public results and activity gates against literal step expectations.</summary>
*)
{endregion}
METHOD PRIVATE CheckResults
FResultsMatch := (FRising.Result = FExpectedResult)
    AND (FFalling.Result = FExpectedResult)
    AND (FDelayedRising.Result = FExpectedDelayedResult)
    AND (FDelayedFalling.Result = FExpectedDelayedResult);
FActivityMatches := (FRising.Enabled = FSubjectEnable)
    AND (FRising.ObservationActive = FExpectedObservation)
    AND (FRising.EvaluationActive = FExpectedEvaluation)
    AND (FFalling.Enabled = FSubjectEnable)
    AND (FFalling.ObservationActive = FExpectedObservation)
    AND (FFalling.EvaluationActive = FExpectedEvaluation)
    AND (FDelayedRising.Enabled = FSubjectEnable)
    AND (FDelayedRising.ObservationActive = FExpectedDelayedObservation)
    AND (FDelayedRising.EvaluationActive = FExpectedDelayedEvaluation)
    AND (FDelayedFalling.Enabled = FSubjectEnable)
    AND (FDelayedFalling.ObservationActive = FExpectedDelayedObservation)
    AND (FDelayedFalling.EvaluationActive = FExpectedDelayedEvaluation);
END_METHOD

{region 'Documentation'}
(*!
<summary>Binds isolated subjects and initializes the outer trace Assertions.</summary>
*)
{endregion}
METHOD PROTECTED Configure
VAR
    Initialized : BOOL;
END_VAR
FPreparationStateCount := 0;
FTestStateCount := 1;
FResetHistory.Initialize(Parent := THIS^,
    AssertionName := 'ResetHistory');
FFirstObservation.Initialize(Parent := THIS^,
    AssertionName := 'FirstObservation');
FHeldFailure.Initialize(Parent := THIS^,
    AssertionName := 'HeldFailure');
FDisabledHistory.Initialize(Parent := THIS^,
    AssertionName := 'DisabledHistory');
FDelayedObservation.Initialize(Parent := THIS^,
    AssertionName := 'DelayedObservation');
FSetupValid := FCapture.Initialize(Buffer := FEvents,
    FifoControl := FCaptureFifo,
    Status := FCaptureStatus);
FRising.BindPublisher(Publisher := FCapture);
Initialized := FRising.Initialize(Parent := THIS^,
    AssertionName := 'Rising',
    ObserveFirstCycle := TRUE);
FSetupValid := FSetupValid AND Initialized;
FFalling.BindPublisher(Publisher := FCapture);
Initialized := FFalling.Initialize(Parent := THIS^,
    AssertionName := 'Falling',
    ObserveFirstCycle := TRUE);
FSetupValid := FSetupValid AND Initialized;
FDelayedRising.BindPublisher(Publisher := FCapture);
Initialized := FDelayedRising.Initialize(Parent := THIS^,
    AssertionName := 'DelayedRising',
    ObserveFirstCycle := FALSE);
FSetupValid := FSetupValid AND Initialized;
FDelayedFalling.BindPublisher(Publisher := FCapture);
Initialized := FDelayedFalling.Initialize(Parent := THIS^,
    AssertionName := 'DelayedFalling',
    ObserveFirstCycle := FALSE);
FSetupValid := FSetupValid AND Initialized;
END_METHOD

{region 'Documentation'}
(*!
<summary>Checks one expected local Failed finding; index is bounded by four subjects.</summary>
*)
{endregion}
METHOD PRIVATE IsFindingValid : BOOL //! TRUE when the selected captured finding satisfies the scenario metadata and diagnostic checks.
VAR_INPUT
    Index : UINT; //! One-based index in the retained isolated event capture.
    ExpectedName : STRING(GVL_Constants.NameLength); //! Independently authored Assertion name expected in the selected finding.
END_VAR
IsFindingValid := (FEvents[Index].SequenceId = UINT_TO_UDINT(Index))
    AND (FEvents[Index].Name = ExpectedName)
    AND (FEvents[Index].OwnerScope = E_OwnerScope.Assertion)
    AND (FEvents[Index].EventType = E_EventType.Result)
    AND (FEvents[Index].State = E_State.Running)
    AND (FEvents[Index].Result = E_Result.Failed)
    AND (FEvents[Index].Message <> '');
END_METHOD

{region 'Documentation'}
(*!
<summary>Completes abort; the trace owns no asynchronous resource.</summary>
*)
{endregion}
METHOD PROTECTED ProcessAbort
VAR_INPUT
    Enable : BOOL; //! Phase permission supplied by the owning Test Case; FALSE does not authorize progression, while observation may continue.
END_VAR
IF Enable THEN
    CompleteAbort();
END_IF;
END_METHOD

{region 'Documentation'}
(*!
<summary>Latches the current trace checkpoint before allowing progression.</summary>
*)
{endregion}
METHOD PROTECTED ProcessAssertions
VAR_INPUT
    Enable : BOOL; //! Phase permission supplied by the owning Test Case; FALSE does not authorize progression, while observation may continue.
END_VAR
VAR
    Check : BOOL;
END_VAR
Check := Enable AND FObservationReady;
FResetHistory(Enable := Check AND (FTrace = TraceResetHistory),
    State := State,
    IN := FStepMatches);
FFirstObservation(Enable := Check AND (FTrace = TraceFirstObservation),
    State := State,
    IN := FStepMatches);
FHeldFailure(Enable := Check AND (FTrace = TraceHeldFailure),
    State := State,
    IN := FStepMatches);
FDisabledHistory(Enable := Check AND (FTrace = TraceDisabledHistory),
    State := State,
    IN := FStepMatches);
FDelayedObservation(Enable := Check AND (FTrace = TraceDelayedObservation),
    State := State,
    IN := FStepMatches);
IF Check THEN
    FChecked := TRUE;
END_IF;
END_METHOD

{region 'Documentation'}
(*!
<summary>No Preparation phase is required.</summary>
*)
{endregion}
METHOD PROTECTED ProcessPreparations
VAR_INPUT
    // SA0033: Required hook; this test has no Preparation phase.
    {attribute 'analysis' := '-33'}
    Enable : BOOL; //! Phase permission supplied by the owning Test Case; FALSE does not authorize progression, while observation may continue.
END_VAR
END_METHOD

{region 'Documentation'}
(*!
<summary>Restarts the trace; subjects consume their reset only with bound inputs.</summary>
*)
{endregion}
METHOD PROTECTED ProcessReset
FStep := StepInitialBoundReset;
FTrace := 0;
FFirstFailedStep := 0;
FChecked := FALSE;
FObservationReady := FALSE;
FStepMatches := TRUE;
FResultsMatch := TRUE;
FActivityMatches := TRUE;
FFindingsMatch := TRUE;
FCapture.Reset();
ResetSubjects();
FResetHistory.Reset();
FFirstObservation.Reset();
FHeldFailure.Reset();
FDisabledHistory.Reset();
FDelayedObservation.Reset();
CompleteReset();
END_METHOD

{region 'Documentation'}
(*!
<summary>Executes one named step per active cycle, after the previous check was latched.</summary>
*)
{endregion}
METHOD PROTECTED ProcessTests
VAR_INPUT
    Enable : BOOL; //! Phase permission supplied by the owning Test Case; FALSE does not authorize progression, while observation may continue.
END_VAR
IF NOT Enable THEN
    RETURN;
END_IF;

IF FChecked THEN
    FChecked := FALSE;
    FObservationReady := FALSE;
    IF FStep = LastStep THEN
        CompleteTests();
        RETURN;
    END_IF;
    FStep := FStep + 1;
END_IF;

IF NOT SelectStep() THEN
    RETURN;
END_IF;
FCapture.Reset();
IF FResetSubjects THEN
    ResetSubjects();
END_IF;
CallSubjects();
CheckResults();
CheckFindings();
FStepMatches := FResultsMatch AND FActivityMatches AND FFindingsMatch;
IF NOT FStepMatches AND (FFirstFailedStep = 0) THEN
    FFirstFailedStep := FStep;
END_IF;
FObservationReady := TRUE;
END_METHOD

{region 'Documentation'}
(*!
<summary>Queues reset without accessing typed cyclic inputs.</summary>
*)
{endregion}
METHOD PRIVATE ResetSubjects
FRising.Reset();
FFalling.Reset();
FDelayedRising.Reset();
FDelayedFalling.Reset();
END_METHOD

